(* PLC project Gaia V6.project, CODESYS CODESYS V3.5 SP22 Patch 2 *)
(* stored: creationDateTime 2026-10-21T15:12:01.6200674, modificationDateTime 2026-10-21T14:27:21.3389871 *)

TYPE DUT_EXC_DOSENSOR : STRUCT
  EXC_OUTPUT_SIGNAL : REAL;  (* [EXC : to other equipment] Dissolved oxygen measure *)
  UPI_INPUT_GLOBAL_LOCAL_FUXA : BOOL;  (* [UPI : functional units to equipment] From UPI_LOCAL_FUXA : global FUXA local active *)
  UPI_INPUT_GLOBAL_LOCAL_HMI : BOOL;  (* From UPI_LOCAL_HMI : global HMI local active *)
  UPI_INPUT_GLOBAL_LOCAL_WEBVISU : BOOL;  (* From UPI_LOCAL_webvisu : global HMI local active *)
END_STRUCT;
END_TYPE

TYPE DUT_INT_DIP1500 : STRUCT
  FUXA_LOCAL_REQUEST : BOOL;  (* [Control mode] From FUXA : local request (pulse or maintained) *)
  FUXA_AUTO_REQUEST : BOOL;  (* From FUXA : auto request, releases the individual FUXA local *)
  HMI_LOCAL_REQUEST : BOOL;  (* From HMI : local request (pulse or maintained) *)
  HMI_AUTO_REQUEST : BOOL;  (* From HMI : auto request, releases the individual HMI local *)
  GLOBAL_LOCAL_FUXA : BOOL;  (* From UPI_LOCAL_FUXA : global FUXA local active *)
  GLOBAL_LOCAL_HMI : BOOL;  (* From UPI_LOCAL_HMI : global HMI local active *)
  LOCAL_FUXA_INDIVIDUAL : BOOL;  (* Memory : individual FUXA local, set by local request, reset by auto request *)
  LOCAL_HMI_INDIVIDUAL : BOOL;  (* Memory : individual HMI local, set by local request, reset by auto request *)
  LOCAL_HMI : BOOL;  (* Result : equipment in HMI local (individual or global), unless WEBVISU local is active *)
  LOCAL_FUXA : BOOL;  (* Result : equipment in FUXA local (individual or global), unless WEBVISU or HMI local is active *)
  AUTO : BOOL;  (* Result : no local mode, commands come from the functional units (UPI) *)
  CMD_RUN : BOOL;  (* [Commands (to pump), from the active source] 0 stop, 1 start *)
  CMD_CLOCKWISE : BOOL;  (* 0 counterclockwise, 1 clockwise *)
  CMD_SAVE_FLASH : BOOL;  (* 1 s pulse to coil 0x0003, saves pump parameters to flash *)
  CMD_VOLUME_MODE : BOOL;  (* 0 time mode, 1 volume mode *)
  CMD_SPEED : REAL;  (* rpm *)
  CMD_MAX_SPEED : REAL;  (* rpm *)
  CMD_RUN_SETPOINT : REAL;  (* ms (time mode) or ml (volume mode), 0 = continuous *)
  CMD_CALIB_COEF : REAL;  (* ml/min or rpm *)
  CMD_FOOT_MODE : WORD;  (* Foot switch input mode *)
  CMD_LEVEL_MODE : WORD;  (* Liquid level input mode *)
  CMD_STATE_OUT_MODE : WORD;  (* State output mode *)
  CMD_ADDRESS : WORD;  (* Modbus address *)
  CMD_BAUD_INDEX : WORD;  (* 0=1200 .. 3=9600 .. 7=115200 *)
  PARAM_WRITE_ENABLE : BOOL;  (* [Parameter writing] 1 = write configuration to the pump, 0 = stop writing *)
  FLASH_SAVE_REQUEST : BOOL;  (* Flash save request (rising edge used) *)
  PARAM_VALID : BOOL;  (* Address 1..31, baud index 0..7, max speed > 0, calibration coefficient > 0 *)
  PULSE_500MS : BOOL;  (* [Write triggers] Square wave, 500 ms period, source of the trigger edges *)
  CMD_CHANGED : BOOL;  (* A command value changed this cycle *)
  CMD_WINDOW : BOOL;  (* Command write window, 3 s after the last change *)
  CMD_TRIGGER : BOOL;  (* Command channel trigger *)
  CONFIG_TRIGGER : BOOL;  (* Configuration channel trigger *)
  PREV_RUN : BOOL;  (* [Previous command values] Previous values for change detection *)
  PREV_CLOCKWISE : BOOL;
  PREV_VOLUME_MODE : BOOL;
  PREV_SAVE_FLASH : BOOL;
  PREV_SPEED : REAL;
  PREV_MAX_SPEED : REAL;
  PREV_RUN_SETPOINT : REAL;
  FBK_FIRMWARE_VERSION : WORD;  (* [Feedback (from pump)] 3+5+8 bits (major+minor+revision) *)
  FBK_HARDWARE_VERSION : WORD;  (* 3+5+8 bits (major+sub+reserved) *)
  FBK_TEMPERATURE : WORD;  (* (raw - 500) / 10 = degC, 65535 = not connected *)
  FBK_LEVEL_ALARM : WORD;  (* 0 no alarm, 1 alarm, 65535 = not connected *)
  FBK_DIGITAL_OUTPUT : WORD;  (* Digital output value *)
  FBK_RUN_ACTUAL : REAL;  (* Current run, ms (time mode) or ml (volume mode) *)
  FBK_RUN_TOTAL : REAL;  (* Accumulated run, ms (time mode) or ml (volume mode) *)
  UDINT_TEMP : UDINT;  (* [Work] Work variable, time mode conversion *)
  WEBVISU_LOCAL_REQUEST : BOOL;  (* From WEBVISU : individual local request *)
  WEBVISU_AUTO_REQUEST : BOOL;  (* From WEBVISU : releases individual WEBVISU local (auto wins) *)
  GLOBAL_LOCAL_WEBVISU : BOOL;  (* From UPI_LOCAL_WEBVISU : global local request *)
  LOCAL_WEBVISU_INDIVIDUAL : BOOL;  (* Memory : individual WEBVISU local request *)
  LOCAL_WEBVISU : BOOL;  (* Effective WEBVISU local : highest source priority *)
  SRC_MAX_MOTOR_SPEED : REAL;  (* [Parameter source] Value typed in the active local supervision *)
  SRC_CALIBRATION_COEFFICIENT : REAL;
  SRC_FOOT_SWITCH_INPUT_MODE : WORD;
  SRC_LIQUID_LEVEL_INPUT_MODE : WORD;
  SRC_STATE_OUTPUT_MODE : WORD;
  SRC_COMMUNICATION_ADDRESS : WORD;
  SRC_BAUD_RATE_INDEX : WORD;
  PREV_SRC_MAX_MOTOR_SPEED : REAL;  (* [Parameter change detection] Previous source values *)
  PREV_SRC_CALIBRATION_COEFFICIENT : REAL;
  PREV_SRC_FOOT_SWITCH_INPUT_MODE : WORD;
  PREV_SRC_LIQUID_LEVEL_INPUT_MODE : WORD;
  PREV_SRC_STATE_OUTPUT_MODE : WORD;
  PREV_SRC_COMMUNICATION_ADDRESS : WORD;
  PREV_SRC_BAUD_RATE_INDEX : WORD;
  PREV_LOCAL_WEBVISU : BOOL;  (* Previous control mode, to ignore the cycle where the source changes *)
  PREV_LOCAL_HMI : BOOL;
  PREV_LOCAL_FUXA : BOOL;
  SOURCE_CHANGED : BOOL;  (* The active local source changed this cycle : no parameter is taken *)
END_STRUCT;
END_TYPE

TYPE DUT_IO_DOSENSOR : STRUCT
  INPUT_SIGNAL : DWORD;  (* [INPUT (field to PLC)] Analog input, raw value *)
  INPUT_SENSOR_FAULT : BOOL;  (* Digital input, sensor fault *)
  OUTPUT_CALIBRATION_HIGH : BOOL;  (* [OUTPUT (PLC to field)] Digital output, high calibration *)
  OUTPUT_CALIBRATION_LOW : BOOL;  (* Digital output, low calibration *)
END_STRUCT;
END_TYPE

TYPE DUT_INT_DOSENSOR : STRUCT
  FUXA_LOCAL_REQUEST : BOOL;  (* [Control mode] From FUXA : local request (pulse or maintained) *)
  FUXA_AUTO_REQUEST : BOOL;  (* From FUXA : auto request, releases the individual FUXA local *)
  HMI_LOCAL_REQUEST : BOOL;  (* From HMI : local request (pulse or maintained) *)
  HMI_AUTO_REQUEST : BOOL;  (* From HMI : auto request, releases the individual HMI local *)
  GLOBAL_LOCAL_FUXA : BOOL;  (* From UPI_LOCAL_FUXA : global FUXA local active *)
  GLOBAL_LOCAL_HMI : BOOL;  (* From UPI_LOCAL_HMI : global HMI local active *)
  LOCAL_FUXA_INDIVIDUAL : BOOL;  (* Memory : individual FUXA local, set by local request, reset by auto request *)
  LOCAL_HMI_INDIVIDUAL : BOOL;  (* Memory : individual HMI local, set by local request, reset by auto request *)
  LOCAL_HMI : BOOL;  (* Result : equipment in HMI local (individual or global), unless WEBVISU local is active *)
  LOCAL_FUXA : BOOL;  (* Result : equipment in FUXA local (individual or global), unless WEBVISU or HMI local is active *)
  WEBVISU_LOCAL_REQUEST : BOOL;  (* From WEBVISU : local request (pulse or maintained) *)
  WEBVISU_AUTO_REQUEST : BOOL;  (* From WEBVISU : auto request, releases the individual WEBVISU local *)
  LOCAL_WEBVISU_INDIVIDUAL : BOOL;  (* Memory : individual WEBVISU local, set by local request, reset by auto request *)
  LOCAL_WEBVISU : BOOL;  (* Result : equipment in WEBVISU local (individual or global), has priority *)
  AUTO : BOOL;  (* Result : no local mode, commands come from the functional units (UPI) *)
  SIGNAL_RAW : DWORD;  (* [Inputs] Raw analog input *)
  FAULT : BOOL;  (* Sensor fault (digital input) *)
  CALIB_HIGH_REQUEST : BOOL;  (* High calibration request from the active source *)
  CALIB_LOW_REQUEST : BOOL;  (* Low calibration request from the active source *)
  SIGNAL : REAL;  (* [Results] Scaled measure *)
  CALIB_HIGH : BOOL;  (* High calibration pulse to sensor (1 s) *)
  CALIB_LOW : BOOL;  (* Low calibration pulse to sensor (1 s) *)
  CALIB_DONE : BOOL;  (* Calibration done message (5 s) *)
  GLOBAL_LOCAL_WEBVISU : BOOL;  (* From UPI_LOCAL_WEBVISU : global local request *)
END_STRUCT;
END_TYPE

TYPE DUT_COM_DOSENSOR : STRUCT
  SCADA_INPUT_CALIBRATION_HIGH : BOOL;  (* [SCADA (FUXA) : input (to PLC)] Coil 1 | DO Calibration High *)
  SCADA_INPUT_CALIBRATION_LOW : BOOL;  (* Coil 2 | DO Calibration Low *)
  SCADA_INPUT_LOCAL_REQUEST : BOOL;  (* Coil 8 | DO Sensor Local Request *)
  SCADA_INPUT_AUTO_REQUEST : BOOL;  (* Coil 9 | DO Sensor Auto Request *)
  SCADA_OUTPUT_FAULT : BOOL;  (* [SCADA (FUXA) : output (from PLC)] DI 10001 | Do sensor fault *)
  SCADA_OUTPUT_CALIBRATION_DONE : BOOL;  (* DI 10002 | Do sensor calibration done *)
  SCADA_OUTPUT_LOCAL_FUXA_ACTIVE : BOOL;  (* DI 10013 | DO Sensor Local FUXA Active *)
  SCADA_OUTPUT_LOCAL_HMI_ACTIVE : BOOL;  (* DI 10014 | DO Sensor Local HMI Active *)
  SCADA_OUTPUT_SIGNAL : DUT_Union_Real_Word;  (* IR 89-90 | DO Sensor Signal *)
  HMI_INPUT_CALIBRATION_HIGH : BOOL;  (* [HMI (local panel, FUXA address + 1000) : input (to PLC)] Coil 1001 | DO Calibration High *)
  HMI_INPUT_CALIBRATION_LOW : BOOL;  (* Coil 1002 | DO Calibration Low *)
  HMI_INPUT_LOCAL_REQUEST : BOOL;  (* Coil 1008 | DO Sensor Local Request *)
  HMI_INPUT_AUTO_REQUEST : BOOL;  (* Coil 1009 | DO Sensor Auto Request *)
  HMI_OUTPUT_FAULT : BOOL;  (* [HMI (local panel, FUXA address + 1000) : output (from PLC)] DI 11001 | Do sensor fault *)
  HMI_OUTPUT_CALIBRATION_DONE : BOOL;  (* DI 11002 | Do sensor calibration done *)
  HMI_OUTPUT_LOCAL_ACTIVE : BOOL;  (* DI 11014 | DO Sensor Local Active *)
  HMI_OUTPUT_SIGNAL : DUT_Union_Real_Word;  (* IR 1089-1090 | DO Sensor Signal *)
  WEBVISU_INPUT_CALIBRATION_HIGH : BOOL;  (* DO Calibration High *)
  WEBVISU_INPUT_CALIBRATION_LOW : BOOL;  (* DO Calibration Low *)
  WEBVISU_INPUT_LOCAL_REQUEST : BOOL;  (* DO Sensor Local Request *)
  WEBVISU_INPUT_AUTO_REQUEST : BOOL;  (* DO Sensor Auto Request *)
  WEBVISU_OUTPUT_FAULT : BOOL;  (* Do sensor fault *)
  WEBVISU_OUTPUT_CALIBRATION_DONE : BOOL;  (* Do sensor calibration done *)
  WEBVISU_OUTPUT_LOCAL_ACTIVE : BOOL;  (* DO Sensor Local Active *)
  WEBVISU_OUTPUT_SIGNAL : DUT_Union_Real_Word;  (* DO Sensor Signal *)
  WEBVISU_OUTPUT_LOCAL_FUXA_ACTIVE : BOOL;  (* Effective FUXA local mode (masked by WEBVISU and HMI priority) *)
  WEBVISU_OUTPUT_LOCAL_HMI_ACTIVE : BOOL;  (* Effective HMI local mode (masked by WEBVISU priority) *)
END_STRUCT;
END_TYPE

TYPE DUT_INT_ADM100W : STRUCT
  FUXA_LOCAL_REQUEST : BOOL;  (* [Control mode] From FUXA : local request (pulse or maintained) *)
  FUXA_AUTO_REQUEST : BOOL;  (* From FUXA : auto request, releases the individual FUXA local *)
  HMI_LOCAL_REQUEST : BOOL;  (* From HMI : local request (pulse or maintained) *)
  HMI_AUTO_REQUEST : BOOL;  (* From HMI : auto request, releases the individual HMI local *)
  GLOBAL_LOCAL_FUXA : BOOL;  (* From UPI_LOCAL_FUXA : global FUXA local active *)
  GLOBAL_LOCAL_HMI : BOOL;  (* From UPI_LOCAL_HMI : global HMI local active *)
  LOCAL_FUXA_INDIVIDUAL : BOOL;  (* Memory : individual FUXA local, set by local request, reset by auto request *)
  LOCAL_HMI_INDIVIDUAL : BOOL;  (* Memory : individual HMI local, set by local request, reset by auto request *)
  LOCAL_HMI : BOOL;  (* Result : equipment in HMI local (individual or global), unless WEBVISU local is active *)
  LOCAL_FUXA : BOOL;  (* Result : equipment in FUXA local (individual or global), unless WEBVISU or HMI local is active *)
  AUTO : BOOL;  (* Result : no local mode, commands come from the functional units (UPI) *)
  ALARM_1 : BOOL;  (* [Alarms] Alarm 1 status *)
  ALARM_2 : BOOL;  (* Alarm 2 status *)
  ALARM_3 : BOOL;  (* Alarm 3 status *)
  ALARM_4 : BOOL;  (* Alarm 4 status *)
  ALARM_5 : BOOL;  (* Alarm 5 status *)
  ALARM_6 : BOOL;  (* Alarm 6 status *)
  ALARM_7 : BOOL;  (* Alarm 7 status *)
  ALARM_8 : BOOL;  (* Alarm 8 status *)
  ALARM_9 : BOOL;  (* Alarm 9 status *)
  ALARM_10 : BOOL;  (* Alarm 10 status *)
  FREQUENCY : REAL;  (* [Measures] Frequency | Hz *)
  L1_L2_VOLTAGE : REAL;  (* L1-L2 Voltage | V *)
  L1_N_VOLTAGE : REAL;  (* L1-N Voltage | V *)
  L1_CURRENT : REAL;  (* L1 Current | A *)
  L1_ACTIVE_POWER : REAL;  (* L1 Active Power | W *)
  L1_APPARENT_POWER : REAL;  (* L1 Apparent Power | VA *)
  L1_REACTIVE_POWER : REAL;  (* L1 Reactive Power | W *)
  L1_CURRENT_PHASE_ANGLE : REAL;  (* L1 Current Phase Angle | deg *)
  L1_POWER_FACTOR : REAL;  (* L1 Power Factor | - *)
  L1_VOLTAGE_THD : REAL;  (* L1 Voltage THD | % *)
  L1_CURRENT_THD : REAL;  (* L1 Current THD | % *)
  L1_MAX_LOAD : REAL;  (* L1 Max Load | % of 60 A *)
  L1_L2_VOLTAGE_PHASE_ANGLE : REAL;  (* L1-L2 Voltage Phase Angle | deg *)
  L2_L3_VOLTAGE : REAL;  (* L2-L3 Voltage | V *)
  L2_N_VOLTAGE : REAL;  (* L2-N Voltage | V *)
  L2_CURRENT : REAL;  (* L2 Current | A *)
  L2_ACTIVE_POWER : REAL;  (* L2 Active Power | W *)
  L2_APPARENT_POWER : REAL;  (* L2 Apparent Power | VA *)
  L2_REACTIVE_POWER : REAL;  (* L2 Reactive Power | W *)
  L2_CURRENT_PHASE_ANGLE : REAL;  (* L2 Current Phase Angle | deg *)
  L2_POWER_FACTOR : REAL;  (* L2 Power Factor | - *)
  L2_VOLTAGE_THD : REAL;  (* L2 Voltage THD | % *)
  L2_CURRENT_THD : REAL;  (* L2 Current THD | % *)
  L2_MAX_LOAD : REAL;  (* L2 Max Load | % of 60 A *)
  L1_L3_VOLTAGE_PHASE_ANGLE : REAL;  (* L1-L3 Voltage Phase Angle | deg *)
  L3_L1_VOLTAGE : REAL;  (* L3-L1 Voltage | V *)
  L3_N_VOLTAGE : REAL;  (* L3-N Voltage | V *)
  L3_CURRENT : REAL;  (* L3 Current | A *)
  L3_ACTIVE_POWER : REAL;  (* L3 Active Power | W *)
  L3_APPARENT_POWER : REAL;  (* L3 Apparent Power | VA *)
  L3_REACTIVE_POWER : REAL;  (* L3 Reactive Power | W *)
  L3_CURRENT_PHASE_ANGLE : REAL;  (* L3 Current Phase Angle | deg *)
  L3_POWER_FACTOR : REAL;  (* L3 Power Factor | - *)
  L3_VOLTAGE_THD : REAL;  (* L3 Voltage THD | % *)
  L3_CURRENT_THD : REAL;  (* L3 Current THD | % *)
  L3_MAX_LOAD : REAL;  (* L3 Max Load | % of 60 A *)
  INTERNAL_TEMPERATURE : REAL;  (* Internal Temperature | degC *)
  ACTIVE_ENERGY : REAL;  (* Active Energy | kWh *)
  APPARENT_ENERGY : REAL;  (* Apparent Energy | per ADM100W config *)
  REACTIVE_ENERGY : REAL;  (* Reactive Energy | kWh *)
  TOTAL_ACTIVE_POWER : REAL;  (* Total Active Power | W *)
  TOTAL_APPARENT_POWER : REAL;  (* Total Apparent Power | VA *)
  TOTAL_REACTIVE_POWER : REAL;  (* Total Reactive Power | W *)
  ALL_PHASE_POWER_FACTOR : REAL;  (* All Phase Power Factor | - *)
  WEBVISU_LOCAL_REQUEST : BOOL;  (* From WEBVISU : individual local request *)
  WEBVISU_AUTO_REQUEST : BOOL;  (* From WEBVISU : releases individual WEBVISU local (auto wins) *)
  GLOBAL_LOCAL_WEBVISU : BOOL;  (* From UPI_LOCAL_WEBVISU : global local request *)
  LOCAL_WEBVISU_INDIVIDUAL : BOOL;  (* Memory : individual WEBVISU local request *)
  LOCAL_WEBVISU : BOOL;  (* Effective WEBVISU local : highest source priority *)
END_STRUCT;
END_TYPE

TYPE DUT_COM_UPI_LOCAL_FUXA : STRUCT
  SCADA_INPUT_LOCAL_REQUEST : BOOL;  (* [SCADA (FUXA) : input (to PLC)] Coil 14 | Global Local FUXA Request *)
  SCADA_INPUT_AUTO_REQUEST : BOOL;  (* Coil 15 | Global Auto FUXA Request *)
  SCADA_OUTPUT_LOCAL_ACTIVE : BOOL;  (* [SCADA (FUXA) : output (from PLC)] DI 10019 | Global Local FUXA Active *)
END_STRUCT;
END_TYPE

TYPE DUT_IO_ADM100W : STRUCT
  SPARE : BOOL;  (* Placeholder, structure not used yet *)
END_STRUCT;
END_TYPE

TYPE DUT_COM_ADM100W : STRUCT
  COM_INPUT_IR : ARRAY[0..87] OF WORD;  (* [COM : Modbus RTU, input (equipment to PLC)] Input registers 0..87, 32-bit float, MSW first (ABCD) *)
  COM_INPUT_COILS : ARRAY[0..1] OF BYTE;  (* Coils 0..9 = alarms 1..10 (byte.bit) *)
  SCADA_INPUT_LOCAL_REQUEST : BOOL;  (* [SCADA (FUXA) : input (to PLC)] Coil 12 | ADM100W Local Request *)
  SCADA_INPUT_AUTO_REQUEST : BOOL;  (* Coil 13 | ADM100W Auto Request *)
  SCADA_OUTPUT_ALARM_1_STATUS : BOOL;  (* [SCADA (FUXA) : output (from PLC)] DI 10003 | ADM100W Alarm 1 Status *)
  SCADA_OUTPUT_ALARM_2_STATUS : BOOL;  (* DI 10004 | ADM100W Alarm 2 Status *)
  SCADA_OUTPUT_ALARM_3_STATUS : BOOL;  (* DI 10005 | ADM100W Alarm 3 Status *)
  SCADA_OUTPUT_ALARM_4_STATUS : BOOL;  (* DI 10006 | ADM100W Alarm 4 Status *)
  SCADA_OUTPUT_ALARM_5_STATUS : BOOL;  (* DI 10007 | ADM100W Alarm 5 Status *)
  SCADA_OUTPUT_ALARM_6_STATUS : BOOL;  (* DI 10008 | ADM100W Alarm 6 Status *)
  SCADA_OUTPUT_ALARM_7_STATUS : BOOL;  (* DI 10009 | ADM100W Alarm 7 Status *)
  SCADA_OUTPUT_ALARM_8_STATUS : BOOL;  (* DI 10010 | ADM100W Alarm 8 Status *)
  SCADA_OUTPUT_ALARM_9_STATUS : BOOL;  (* DI 10011 | ADM100W Alarm 9 Status *)
  SCADA_OUTPUT_ALARM_10_STATUS : BOOL;  (* DI 10012 | ADM100W Alarm 10 Status *)
  SCADA_OUTPUT_LOCAL_FUXA_ACTIVE : BOOL;  (* DI 10017 | ADM100W Local FUXA Active *)
  SCADA_OUTPUT_LOCAL_HMI_ACTIVE : BOOL;  (* DI 10018 | ADM100W Local HMI Active *)
  SCADA_OUTPUT_FREQUENCY : DUT_Union_Real_Word;  (* IR 1-2 | ADM100W Frequency | Hz *)
  SCADA_OUTPUT_L1_L2_VOLTAGE : DUT_Union_Real_Word;  (* IR 3-4 | ADM100W L1-L2 Voltage | V *)
  SCADA_OUTPUT_L1_N_VOLTAGE : DUT_Union_Real_Word;  (* IR 5-6 | ADM100W L1-N Voltage | V *)
  SCADA_OUTPUT_L1_CURRENT : DUT_Union_Real_Word;  (* IR 7-8 | ADM100W L1 Current | A *)
  SCADA_OUTPUT_L1_ACTIVE_POWER : DUT_Union_Real_Word;  (* IR 9-10 | ADM100W L1 Active Power *)
  SCADA_OUTPUT_L1_APPARENT_POWER : DUT_Union_Real_Word;  (* IR 11-12 | ADM100W L1 Apparent Power *)
  SCADA_OUTPUT_L1_REACTIVE_POWER : DUT_Union_Real_Word;  (* IR 13-14 | ADM100W L1 Reactive Power *)
  SCADA_OUTPUT_L1_CURRENT_PHASE_ANGLE : DUT_Union_Real_Word;  (* IR 15-16 | ADM100W L1 Current Phase Angle | deg *)
  SCADA_OUTPUT_L1_POWER_FACTOR : DUT_Union_Real_Word;  (* IR 17-18 | ADM100W L1 Power Factor *)
  SCADA_OUTPUT_L1_VOLTAGE_THD : DUT_Union_Real_Word;  (* IR 19-20 | ADM100W L1 Voltage THD | % *)
  SCADA_OUTPUT_L1_CURRENT_THD : DUT_Union_Real_Word;  (* IR 21-22 | ADM100W L1 Current THD | % *)
  SCADA_OUTPUT_L1_MAX_LOAD : DUT_Union_Real_Word;  (* IR 23-24 | ADM100W L1 Max Load *)
  SCADA_OUTPUT_L1_L2_VOLTAGE_PHASE_ANGLE : DUT_Union_Real_Word;  (* IR 25-26 | ADM100W L1-L2 Voltage Phase Angle | deg *)
  SCADA_OUTPUT_L2_L3_VOLTAGE : DUT_Union_Real_Word;  (* IR 27-28 | ADM100W L2-L3 Voltage | V *)
  SCADA_OUTPUT_L2_N_VOLTAGE : DUT_Union_Real_Word;  (* IR 29-30 | ADM100W L2-N Voltage | V *)
  SCADA_OUTPUT_L2_CURRENT : DUT_Union_Real_Word;  (* IR 31-32 | ADM100W L2 Current | A *)
  SCADA_OUTPUT_L2_ACTIVE_POWER : DUT_Union_Real_Word;  (* IR 33-34 | ADM100W L2 Active Power *)
  SCADA_OUTPUT_L2_APPARENT_POWER : DUT_Union_Real_Word;  (* IR 35-36 | ADM100W L2 Apparent Power *)
  SCADA_OUTPUT_L2_REACTIVE_POWER : DUT_Union_Real_Word;  (* IR 37-38 | ADM100W L2 Reactive Power *)
  SCADA_OUTPUT_L2_CURRENT_PHASE_ANGLE : DUT_Union_Real_Word;  (* IR 39-40 | ADM100W L2 Current Phase Angle | deg *)
  SCADA_OUTPUT_L2_POWER_FACTOR : DUT_Union_Real_Word;  (* IR 41-42 | ADM100W L2 Power Factor *)
  SCADA_OUTPUT_L2_VOLTAGE_THD : DUT_Union_Real_Word;  (* IR 43-44 | ADM100W L2 Voltage THD | % *)
  SCADA_OUTPUT_L2_CURRENT_THD : DUT_Union_Real_Word;  (* IR 45-46 | ADM100W L2 Current THD | % *)
  SCADA_OUTPUT_L2_MAX_LOAD : DUT_Union_Real_Word;  (* IR 47-48 | ADM100W L2 Max Load *)
  SCADA_OUTPUT_L1_L3_VOLTAGE_PHASE_ANGLE : DUT_Union_Real_Word;  (* IR 49-50 | ADM100W L1-L3 Voltage Phase Angle | deg *)
  SCADA_OUTPUT_L3_L1_VOLTAGE : DUT_Union_Real_Word;  (* IR 51-52 | ADM100W L3-L1 Voltage | V *)
  SCADA_OUTPUT_L3_N_VOLTAGE : DUT_Union_Real_Word;  (* IR 53-54 | ADM100W L3-N Voltage | V *)
  SCADA_OUTPUT_L3_CURRENT : DUT_Union_Real_Word;  (* IR 55-56 | ADM100W L3 Current | A *)
  SCADA_OUTPUT_L3_ACTIVE_POWER : DUT_Union_Real_Word;  (* IR 57-58 | ADM100W L3 Active Power *)
  SCADA_OUTPUT_L3_APPARENT_POWER : DUT_Union_Real_Word;  (* IR 59-60 | ADM100W L3 Apparent Power *)
  SCADA_OUTPUT_L3_REACTIVE_POWER : DUT_Union_Real_Word;  (* IR 61-62 | ADM100W L3 Reactive Power *)
  SCADA_OUTPUT_L3_CURRENT_PHASE_ANGLE : DUT_Union_Real_Word;  (* IR 63-64 | ADM100W L3 Current Phase Angle | deg *)
  SCADA_OUTPUT_L3_POWER_FACTOR : DUT_Union_Real_Word;  (* IR 65-66 | ADM100W L3 Power Factor *)
  SCADA_OUTPUT_L3_VOLTAGE_THD : DUT_Union_Real_Word;  (* IR 67-68 | ADM100W L3 Voltage THD | % *)
  SCADA_OUTPUT_L3_CURRENT_THD : DUT_Union_Real_Word;  (* IR 69-70 | ADM100W L3 Current THD | % *)
  SCADA_OUTPUT_L3_MAX_LOAD : DUT_Union_Real_Word;  (* IR 71-72 | ADM100W L3 Max Load *)
  SCADA_OUTPUT_INTERNAL_TEMPERATURE : DUT_Union_Real_Word;  (* IR 73-74 | ADM100W Internal Temperature *)
  SCADA_OUTPUT_ACTIVE_ENERGY : DUT_Union_Real_Word;  (* IR 75-76 | ADM100W Active Energy *)
  SCADA_OUTPUT_APPARENT_ENERGY : DUT_Union_Real_Word;  (* IR 77-78 | ADM100W Apparent Energy *)
  SCADA_OUTPUT_REACTIVE_ENERGY : DUT_Union_Real_Word;  (* IR 79-80 | ADM100W Reactive Energy *)
  SCADA_OUTPUT_TOTAL_ACTIVE_POWER : DUT_Union_Real_Word;  (* IR 81-82 | ADM100W Total Active Power *)
  SCADA_OUTPUT_TOTAL_APPARENT_POWER : DUT_Union_Real_Word;  (* IR 83-84 | ADM100W Total Apparent Power *)
  SCADA_OUTPUT_TOTAL_REACTIVE_POWER : DUT_Union_Real_Word;  (* IR 85-86 | ADM100W Total Reactive Power *)
  SCADA_OUTPUT_ALL_PHASE_POWER_FACTOR : DUT_Union_Real_Word;  (* IR 87-88 | ADM100W All Phase Power Factor *)
  HMI_INPUT_LOCAL_REQUEST : BOOL;  (* [HMI (local panel, FUXA address + 1000) : input (to PLC)] Coil 1012 | ADM100W Local Request *)
  HMI_INPUT_AUTO_REQUEST : BOOL;  (* Coil 1013 | ADM100W Auto Request *)
  HMI_OUTPUT_ALARM_1_STATUS : BOOL;  (* [HMI (local panel, FUXA address + 1000) : output (from PLC)] DI 11003 | ADM100W Alarm 1 Status *)
  HMI_OUTPUT_ALARM_2_STATUS : BOOL;  (* DI 11004 | ADM100W Alarm 2 Status *)
  HMI_OUTPUT_ALARM_3_STATUS : BOOL;  (* DI 11005 | ADM100W Alarm 3 Status *)
  HMI_OUTPUT_ALARM_4_STATUS : BOOL;  (* DI 11006 | ADM100W Alarm 4 Status *)
  HMI_OUTPUT_ALARM_5_STATUS : BOOL;  (* DI 11007 | ADM100W Alarm 5 Status *)
  HMI_OUTPUT_ALARM_6_STATUS : BOOL;  (* DI 11008 | ADM100W Alarm 6 Status *)
  HMI_OUTPUT_ALARM_7_STATUS : BOOL;  (* DI 11009 | ADM100W Alarm 7 Status *)
  HMI_OUTPUT_ALARM_8_STATUS : BOOL;  (* DI 11010 | ADM100W Alarm 8 Status *)
  HMI_OUTPUT_ALARM_9_STATUS : BOOL;  (* DI 11011 | ADM100W Alarm 9 Status *)
  HMI_OUTPUT_ALARM_10_STATUS : BOOL;  (* DI 11012 | ADM100W Alarm 10 Status *)
  HMI_OUTPUT_LOCAL_ACTIVE : BOOL;  (* DI 11018 | ADM100W Local Active *)
  HMI_OUTPUT_FREQUENCY : DUT_Union_Real_Word;  (* IR 1001-1002 | ADM100W Frequency | Hz *)
  HMI_OUTPUT_L1_L2_VOLTAGE : DUT_Union_Real_Word;  (* IR 1003-1004 | ADM100W L1-L2 Voltage | V *)
  HMI_OUTPUT_L1_N_VOLTAGE : DUT_Union_Real_Word;  (* IR 1005-1006 | ADM100W L1-N Voltage | V *)
  HMI_OUTPUT_L1_CURRENT : DUT_Union_Real_Word;  (* IR 1007-1008 | ADM100W L1 Current | A *)
  HMI_OUTPUT_L1_ACTIVE_POWER : DUT_Union_Real_Word;  (* IR 1009-1010 | ADM100W L1 Active Power *)
  HMI_OUTPUT_L1_APPARENT_POWER : DUT_Union_Real_Word;  (* IR 1011-1012 | ADM100W L1 Apparent Power *)
  HMI_OUTPUT_L1_REACTIVE_POWER : DUT_Union_Real_Word;  (* IR 1013-1014 | ADM100W L1 Reactive Power *)
  HMI_OUTPUT_L1_CURRENT_PHASE_ANGLE : DUT_Union_Real_Word;  (* IR 1015-1016 | ADM100W L1 Current Phase Angle | deg *)
  HMI_OUTPUT_L1_POWER_FACTOR : DUT_Union_Real_Word;  (* IR 1017-1018 | ADM100W L1 Power Factor *)
  HMI_OUTPUT_L1_VOLTAGE_THD : DUT_Union_Real_Word;  (* IR 1019-1020 | ADM100W L1 Voltage THD | % *)
  HMI_OUTPUT_L1_CURRENT_THD : DUT_Union_Real_Word;  (* IR 1021-1022 | ADM100W L1 Current THD | % *)
  HMI_OUTPUT_L1_MAX_LOAD : DUT_Union_Real_Word;  (* IR 1023-1024 | ADM100W L1 Max Load *)
  HMI_OUTPUT_L1_L2_VOLTAGE_PHASE_ANGLE : DUT_Union_Real_Word;  (* IR 1025-1026 | ADM100W L1-L2 Voltage Phase Angle | deg *)
  HMI_OUTPUT_L2_L3_VOLTAGE : DUT_Union_Real_Word;  (* IR 1027-1028 | ADM100W L2-L3 Voltage | V *)
  HMI_OUTPUT_L2_N_VOLTAGE : DUT_Union_Real_Word;  (* IR 1029-1030 | ADM100W L2-N Voltage | V *)
  HMI_OUTPUT_L2_CURRENT : DUT_Union_Real_Word;  (* IR 1031-1032 | ADM100W L2 Current | A *)
  HMI_OUTPUT_L2_ACTIVE_POWER : DUT_Union_Real_Word;  (* IR 1033-1034 | ADM100W L2 Active Power *)
  HMI_OUTPUT_L2_APPARENT_POWER : DUT_Union_Real_Word;  (* IR 1035-1036 | ADM100W L2 Apparent Power *)
  HMI_OUTPUT_L2_REACTIVE_POWER : DUT_Union_Real_Word;  (* IR 1037-1038 | ADM100W L2 Reactive Power *)
  HMI_OUTPUT_L2_CURRENT_PHASE_ANGLE : DUT_Union_Real_Word;  (* IR 1039-1040 | ADM100W L2 Current Phase Angle | deg *)
  HMI_OUTPUT_L2_POWER_FACTOR : DUT_Union_Real_Word;  (* IR 1041-1042 | ADM100W L2 Power Factor *)
  HMI_OUTPUT_L2_VOLTAGE_THD : DUT_Union_Real_Word;  (* IR 1043-1044 | ADM100W L2 Voltage THD | % *)
  HMI_OUTPUT_L2_CURRENT_THD : DUT_Union_Real_Word;  (* IR 1045-1046 | ADM100W L2 Current THD | % *)
  HMI_OUTPUT_L2_MAX_LOAD : DUT_Union_Real_Word;  (* IR 1047-1048 | ADM100W L2 Max Load *)
  HMI_OUTPUT_L1_L3_VOLTAGE_PHASE_ANGLE : DUT_Union_Real_Word;  (* IR 1049-1050 | ADM100W L1-L3 Voltage Phase Angle | deg *)
  HMI_OUTPUT_L3_L1_VOLTAGE : DUT_Union_Real_Word;  (* IR 1051-1052 | ADM100W L3-L1 Voltage | V *)
  HMI_OUTPUT_L3_N_VOLTAGE : DUT_Union_Real_Word;  (* IR 1053-1054 | ADM100W L3-N Voltage | V *)
  HMI_OUTPUT_L3_CURRENT : DUT_Union_Real_Word;  (* IR 1055-1056 | ADM100W L3 Current | A *)
  HMI_OUTPUT_L3_ACTIVE_POWER : DUT_Union_Real_Word;  (* IR 1057-1058 | ADM100W L3 Active Power *)
  HMI_OUTPUT_L3_APPARENT_POWER : DUT_Union_Real_Word;  (* IR 1059-1060 | ADM100W L3 Apparent Power *)
  HMI_OUTPUT_L3_REACTIVE_POWER : DUT_Union_Real_Word;  (* IR 1061-1062 | ADM100W L3 Reactive Power *)
  HMI_OUTPUT_L3_CURRENT_PHASE_ANGLE : DUT_Union_Real_Word;  (* IR 1063-1064 | ADM100W L3 Current Phase Angle | deg *)
  HMI_OUTPUT_L3_POWER_FACTOR : DUT_Union_Real_Word;  (* IR 1065-1066 | ADM100W L3 Power Factor *)
  HMI_OUTPUT_L3_VOLTAGE_THD : DUT_Union_Real_Word;  (* IR 1067-1068 | ADM100W L3 Voltage THD | % *)
  HMI_OUTPUT_L3_CURRENT_THD : DUT_Union_Real_Word;  (* IR 1069-1070 | ADM100W L3 Current THD | % *)
  HMI_OUTPUT_L3_MAX_LOAD : DUT_Union_Real_Word;  (* IR 1071-1072 | ADM100W L3 Max Load *)
  HMI_OUTPUT_INTERNAL_TEMPERATURE : DUT_Union_Real_Word;  (* IR 1073-1074 | ADM100W Internal Temperature *)
  HMI_OUTPUT_ACTIVE_ENERGY : DUT_Union_Real_Word;  (* IR 1075-1076 | ADM100W Active Energy *)
  HMI_OUTPUT_APPARENT_ENERGY : DUT_Union_Real_Word;  (* IR 1077-1078 | ADM100W Apparent Energy *)
  HMI_OUTPUT_REACTIVE_ENERGY : DUT_Union_Real_Word;  (* IR 1079-1080 | ADM100W Reactive Energy *)
  HMI_OUTPUT_TOTAL_ACTIVE_POWER : DUT_Union_Real_Word;  (* IR 1081-1082 | ADM100W Total Active Power *)
  HMI_OUTPUT_TOTAL_APPARENT_POWER : DUT_Union_Real_Word;  (* IR 1083-1084 | ADM100W Total Apparent Power *)
  HMI_OUTPUT_TOTAL_REACTIVE_POWER : DUT_Union_Real_Word;  (* IR 1085-1086 | ADM100W Total Reactive Power *)
  HMI_OUTPUT_ALL_PHASE_POWER_FACTOR : DUT_Union_Real_Word;  (* IR 1087-1088 | ADM100W All Phase Power Factor *)
  WEBVISU_INPUT_LOCAL_REQUEST : BOOL;  (* [WEBVISU : direct IEC variable] ADM100W Local Request *)
  WEBVISU_INPUT_AUTO_REQUEST : BOOL;  (* [WEBVISU : direct IEC variable] ADM100W Auto Request *)
  WEBVISU_OUTPUT_ALARM_1_STATUS : BOOL;  (* [WEBVISU : direct IEC variable] ADM100W Alarm 1 Status *)
  WEBVISU_OUTPUT_ALARM_2_STATUS : BOOL;  (* [WEBVISU : direct IEC variable] ADM100W Alarm 2 Status *)
  WEBVISU_OUTPUT_ALARM_3_STATUS : BOOL;  (* [WEBVISU : direct IEC variable] ADM100W Alarm 3 Status *)
  WEBVISU_OUTPUT_ALARM_4_STATUS : BOOL;  (* [WEBVISU : direct IEC variable] ADM100W Alarm 4 Status *)
  WEBVISU_OUTPUT_ALARM_5_STATUS : BOOL;  (* [WEBVISU : direct IEC variable] ADM100W Alarm 5 Status *)
  WEBVISU_OUTPUT_ALARM_6_STATUS : BOOL;  (* [WEBVISU : direct IEC variable] ADM100W Alarm 6 Status *)
  WEBVISU_OUTPUT_ALARM_7_STATUS : BOOL;  (* [WEBVISU : direct IEC variable] ADM100W Alarm 7 Status *)
  WEBVISU_OUTPUT_ALARM_8_STATUS : BOOL;  (* [WEBVISU : direct IEC variable] ADM100W Alarm 8 Status *)
  WEBVISU_OUTPUT_ALARM_9_STATUS : BOOL;  (* [WEBVISU : direct IEC variable] ADM100W Alarm 9 Status *)
  WEBVISU_OUTPUT_ALARM_10_STATUS : BOOL;  (* [WEBVISU : direct IEC variable] ADM100W Alarm 10 Status *)
  WEBVISU_OUTPUT_LOCAL_ACTIVE : BOOL;  (* [WEBVISU : direct IEC variable] ADM100W Local Active *)
  WEBVISU_OUTPUT_FREQUENCY : DUT_Union_Real_Word;  (* [WEBVISU : direct IEC variable] ADM100W Frequency | Hz *)
  WEBVISU_OUTPUT_L1_L2_VOLTAGE : DUT_Union_Real_Word;  (* [WEBVISU : direct IEC variable] ADM100W L1-L2 Voltage | V *)
  WEBVISU_OUTPUT_L1_N_VOLTAGE : DUT_Union_Real_Word;  (* [WEBVISU : direct IEC variable] ADM100W L1-N Voltage | V *)
  WEBVISU_OUTPUT_L1_CURRENT : DUT_Union_Real_Word;  (* [WEBVISU : direct IEC variable] ADM100W L1 Current | A *)
  WEBVISU_OUTPUT_L1_ACTIVE_POWER : DUT_Union_Real_Word;  (* [WEBVISU : direct IEC variable] ADM100W L1 Active Power *)
  WEBVISU_OUTPUT_L1_APPARENT_POWER : DUT_Union_Real_Word;  (* [WEBVISU : direct IEC variable] ADM100W L1 Apparent Power *)
  WEBVISU_OUTPUT_L1_REACTIVE_POWER : DUT_Union_Real_Word;  (* [WEBVISU : direct IEC variable] ADM100W L1 Reactive Power *)
  WEBVISU_OUTPUT_L1_CURRENT_PHASE_ANGLE : DUT_Union_Real_Word;  (* [WEBVISU : direct IEC variable] ADM100W L1 Current Phase Angle | deg *)
  WEBVISU_OUTPUT_L1_POWER_FACTOR : DUT_Union_Real_Word;  (* [WEBVISU : direct IEC variable] ADM100W L1 Power Factor *)
  WEBVISU_OUTPUT_L1_VOLTAGE_THD : DUT_Union_Real_Word;  (* [WEBVISU : direct IEC variable] ADM100W L1 Voltage THD | % *)
  WEBVISU_OUTPUT_L1_CURRENT_THD : DUT_Union_Real_Word;  (* [WEBVISU : direct IEC variable] ADM100W L1 Current THD | % *)
  WEBVISU_OUTPUT_L1_MAX_LOAD : DUT_Union_Real_Word;  (* [WEBVISU : direct IEC variable] ADM100W L1 Max Load *)
  WEBVISU_OUTPUT_L1_L2_VOLTAGE_PHASE_ANGLE : DUT_Union_Real_Word;  (* [WEBVISU : direct IEC variable] ADM100W L1-L2 Voltage Phase Angle | deg *)
  WEBVISU_OUTPUT_L2_L3_VOLTAGE : DUT_Union_Real_Word;  (* [WEBVISU : direct IEC variable] ADM100W L2-L3 Voltage | V *)
  WEBVISU_OUTPUT_L2_N_VOLTAGE : DUT_Union_Real_Word;  (* [WEBVISU : direct IEC variable] ADM100W L2-N Voltage | V *)
  WEBVISU_OUTPUT_L2_CURRENT : DUT_Union_Real_Word;  (* [WEBVISU : direct IEC variable] ADM100W L2 Current | A *)
  WEBVISU_OUTPUT_L2_ACTIVE_POWER : DUT_Union_Real_Word;  (* [WEBVISU : direct IEC variable] ADM100W L2 Active Power *)
  WEBVISU_OUTPUT_L2_APPARENT_POWER : DUT_Union_Real_Word;  (* [WEBVISU : direct IEC variable] ADM100W L2 Apparent Power *)
  WEBVISU_OUTPUT_L2_REACTIVE_POWER : DUT_Union_Real_Word;  (* [WEBVISU : direct IEC variable] ADM100W L2 Reactive Power *)
  WEBVISU_OUTPUT_L2_CURRENT_PHASE_ANGLE : DUT_Union_Real_Word;  (* [WEBVISU : direct IEC variable] ADM100W L2 Current Phase Angle | deg *)
  WEBVISU_OUTPUT_L2_POWER_FACTOR : DUT_Union_Real_Word;  (* [WEBVISU : direct IEC variable] ADM100W L2 Power Factor *)
  WEBVISU_OUTPUT_L2_VOLTAGE_THD : DUT_Union_Real_Word;  (* [WEBVISU : direct IEC variable] ADM100W L2 Voltage THD | % *)
  WEBVISU_OUTPUT_L2_CURRENT_THD : DUT_Union_Real_Word;  (* [WEBVISU : direct IEC variable] ADM100W L2 Current THD | % *)
  WEBVISU_OUTPUT_L2_MAX_LOAD : DUT_Union_Real_Word;  (* [WEBVISU : direct IEC variable] ADM100W L2 Max Load *)
  WEBVISU_OUTPUT_L1_L3_VOLTAGE_PHASE_ANGLE : DUT_Union_Real_Word;  (* [WEBVISU : direct IEC variable] ADM100W L1-L3 Voltage Phase Angle | deg *)
  WEBVISU_OUTPUT_L3_L1_VOLTAGE : DUT_Union_Real_Word;  (* [WEBVISU : direct IEC variable] ADM100W L3-L1 Voltage | V *)
  WEBVISU_OUTPUT_L3_N_VOLTAGE : DUT_Union_Real_Word;  (* [WEBVISU : direct IEC variable] ADM100W L3-N Voltage | V *)
  WEBVISU_OUTPUT_L3_CURRENT : DUT_Union_Real_Word;  (* [WEBVISU : direct IEC variable] ADM100W L3 Current | A *)
  WEBVISU_OUTPUT_L3_ACTIVE_POWER : DUT_Union_Real_Word;  (* [WEBVISU : direct IEC variable] ADM100W L3 Active Power *)
  WEBVISU_OUTPUT_L3_APPARENT_POWER : DUT_Union_Real_Word;  (* [WEBVISU : direct IEC variable] ADM100W L3 Apparent Power *)
  WEBVISU_OUTPUT_L3_REACTIVE_POWER : DUT_Union_Real_Word;  (* [WEBVISU : direct IEC variable] ADM100W L3 Reactive Power *)
  WEBVISU_OUTPUT_L3_CURRENT_PHASE_ANGLE : DUT_Union_Real_Word;  (* [WEBVISU : direct IEC variable] ADM100W L3 Current Phase Angle | deg *)
  WEBVISU_OUTPUT_L3_POWER_FACTOR : DUT_Union_Real_Word;  (* [WEBVISU : direct IEC variable] ADM100W L3 Power Factor *)
  WEBVISU_OUTPUT_L3_VOLTAGE_THD : DUT_Union_Real_Word;  (* [WEBVISU : direct IEC variable] ADM100W L3 Voltage THD | % *)
  WEBVISU_OUTPUT_L3_CURRENT_THD : DUT_Union_Real_Word;  (* [WEBVISU : direct IEC variable] ADM100W L3 Current THD | % *)
  WEBVISU_OUTPUT_L3_MAX_LOAD : DUT_Union_Real_Word;  (* [WEBVISU : direct IEC variable] ADM100W L3 Max Load *)
  WEBVISU_OUTPUT_INTERNAL_TEMPERATURE : DUT_Union_Real_Word;  (* [WEBVISU : direct IEC variable] ADM100W Internal Temperature *)
  WEBVISU_OUTPUT_ACTIVE_ENERGY : DUT_Union_Real_Word;  (* [WEBVISU : direct IEC variable] ADM100W Active Energy *)
  WEBVISU_OUTPUT_APPARENT_ENERGY : DUT_Union_Real_Word;  (* [WEBVISU : direct IEC variable] ADM100W Apparent Energy *)
  WEBVISU_OUTPUT_REACTIVE_ENERGY : DUT_Union_Real_Word;  (* [WEBVISU : direct IEC variable] ADM100W Reactive Energy *)
  WEBVISU_OUTPUT_TOTAL_ACTIVE_POWER : DUT_Union_Real_Word;  (* [WEBVISU : direct IEC variable] ADM100W Total Active Power *)
  WEBVISU_OUTPUT_TOTAL_APPARENT_POWER : DUT_Union_Real_Word;  (* [WEBVISU : direct IEC variable] ADM100W Total Apparent Power *)
  WEBVISU_OUTPUT_TOTAL_REACTIVE_POWER : DUT_Union_Real_Word;  (* [WEBVISU : direct IEC variable] ADM100W Total Reactive Power *)
  WEBVISU_OUTPUT_ALL_PHASE_POWER_FACTOR : DUT_Union_Real_Word;  (* [WEBVISU : direct IEC variable] ADM100W All Phase Power Factor *)
  WEBVISU_OUTPUT_LOCAL_FUXA_ACTIVE : BOOL;  (* Effective FUXA local mode (masked by WEBVISU and HMI priority) *)
  WEBVISU_OUTPUT_LOCAL_HMI_ACTIVE : BOOL;  (* Effective HMI local mode (masked by WEBVISU priority) *)
END_STRUCT;
END_TYPE

TYPE DUT_EXC_ADM100W : STRUCT
  EXC_OUTPUT_FREQUENCY : REAL;  (* [EXC : to other equipment] Hz *)
  EXC_OUTPUT_L1_N_VOLTAGE : REAL;  (* V *)
  EXC_OUTPUT_L1_CURRENT : REAL;  (* A *)
  EXC_OUTPUT_L1_ACTIVE_POWER : REAL;  (* W *)
  EXC_OUTPUT_L1_APPARENT_POWER : REAL;  (* VA *)
  EXC_OUTPUT_L1_REACTIVE_POWER : REAL;  (* VAr *)
  EXC_OUTPUT_L1_POWER_FACTOR : REAL;  (* - *)
  EXC_OUTPUT_L1_VOLTAGE_THD : REAL;  (* % *)
  EXC_OUTPUT_L1_CURRENT_THD : REAL;  (* % *)
  EXC_OUTPUT_L1_MAX_LOAD : REAL;  (* % of 60 A *)
  EXC_OUTPUT_INTERNAL_TEMPERATURE : REAL;  (* degC *)
  EXC_OUTPUT_ACTIVE_ENERGY : REAL;  (* kWh *)
  EXC_OUTPUT_DATA_VALID : BOOL;  (* FALSE = values not usable. Not managed yet (no Modbus diagnostic) *)
  UPI_INPUT_GLOBAL_LOCAL_FUXA : BOOL;  (* [UPI : functional units to equipment] From UPI_LOCAL_FUXA : global FUXA local active *)
  UPI_INPUT_GLOBAL_LOCAL_HMI : BOOL;  (* From UPI_LOCAL_HMI : global HMI local active *)
  UPI_INPUT_GLOBAL_LOCAL_WEBVISU : BOOL;  (* From UPI_LOCAL_WEBVISU : global WEBVISU local active *)
END_STRUCT;
END_TYPE

TYPE DUT_COM_DIP1500 : STRUCT
  COM_INPUT_IR : ARRAY[0..4] OF WORD;  (* [COM : Modbus RTU, input (equipment to PLC)] Input registers 0x3001..0x3005 *)
  COM_INPUT_HR_COUNTERS : ARRAY[0..3] OF WORD;  (* Holding registers 0x4007..0x400A (read) *)
  COM_OUTPUT_COILS : ARRAY[0..3] OF BOOL;  (* [COM : Modbus RTU, output (PLC to equipment)] Coils 0x0001..0x0004 *)
  COM_OUTPUT_HR_CMD : ARRAY[0..5] OF WORD;  (* Holding registers 0x4001..0x4006 (write) *)
  COM_OUTPUT_HR_CONFIG : ARRAY[0..6] OF WORD;  (* Holding registers 0x400B..0x4011 (write) *)
  COM_OUTPUT_CMD_TRIGGER : BOOL;  (* Rising edge trigger of the command write channel(s), mapped in the Modbus slave I/O mapping *)
  COM_OUTPUT_CONFIG_TRIGGER : BOOL;  (* Rising edge trigger of the configuration write channel, mapped in the Modbus slave I/O mapping *)
  SCADA_INPUT_MOTOR_START_STOP : BOOL;  (* [SCADA (FUXA) : input (to PLC)] Coil 3 | DIP1500 Motor Start Stop *)
  SCADA_INPUT_MOTOR_DIRECTION : BOOL;  (* Coil 4 | DIP1500 Motor Direction *)
  SCADA_INPUT_FLASH_SAVE : BOOL;  (* Coil 5 | DIP1500 Flash Save *)
  SCADA_INPUT_OPERATION_MODE : BOOL;  (* Coil 6 | DIP1500 Operation Mode *)
  SCADA_INPUT_PARAM_WRITE_ENABLE : BOOL;  (* Coil 7 | DIP1500 Parameter Write Enable *)
  SCADA_INPUT_LOCAL_REQUEST : BOOL;  (* Coil 10 | DIP1500 Local Request *)
  SCADA_INPUT_AUTO_REQUEST : BOOL;  (* Coil 11 | DIP1500 Auto Request *)
  SCADA_INPUT_FOOT_SWITCH_INPUT_MODE : WORD;  (* HR 9 | DIP1500 Foot Switch Input Mode *)
  SCADA_INPUT_LIQUID_LEVEL_INPUT_MODE : WORD;  (* HR 10 | DIP1500 Liquid Level Input Mode *)
  SCADA_INPUT_STATE_OUTPUT_MODE : WORD;  (* HR 11 | DIP1500 State Output Mode *)
  SCADA_INPUT_COMMUNICATION_ADDRESS : WORD;  (* HR 12 | DIP1500 Communication Address *)
  SCADA_INPUT_BAUD_RATE_INDEX : WORD;  (* HR 13 | DIP1500 Baud Rate Index | index *)
  SCADA_INPUT_MOTOR_SPEED : DUT_Union_Real_Word;  (* HR 1-2 | DIP1500 Motor Speed | rpm *)
  SCADA_INPUT_MAX_MOTOR_SPEED : DUT_Union_Real_Word;  (* HR 3-4 | DIP1500 Max Motor Speed | rpm *)
  SCADA_INPUT_RUN_TIME_OR_VOLUME_SETPOINT : DUT_Union_Real_Word;  (* HR 5-6 | DIP1500 Run Time Or Volume Setpoint | ms (time mode) / ml (volume mode) *)
  SCADA_INPUT_FLOW_RATE_OR_SPEED_CALIBRATION_COEFFICIENT : DUT_Union_Real_Word;  (* HR 7-8 | DIP1500 Flow Rate Or Speed Calibration Coefficient | ml/min or rpm *)
  SCADA_OUTPUT_LOCAL_FUXA_ACTIVE : BOOL;  (* [SCADA (FUXA) : output (from PLC)] DI 10015 | DIP1500 Local FUXA Active *)
  SCADA_OUTPUT_LOCAL_HMI_ACTIVE : BOOL;  (* DI 10016 | DIP1500 Local HMI Active *)
  SCADA_OUTPUT_FIRMWARE_VERSION : WORD;  (* IR 91 | DIP1500 Firmware Version | 3+5+8 bits (major+minor+revision) *)
  SCADA_OUTPUT_HARDWARE_VERSION : WORD;  (* IR 92 | DIP1500 Hardware Version | 3+5+8 bits (major+minor+revision) *)
  SCADA_OUTPUT_TEMPERATURE : WORD;  (* IR 93 | DIP1500 Temperature | degC | (raw - 500) / 10 *)
  SCADA_OUTPUT_FLOAT_LEVEL_ALARM : WORD;  (* IR 94 | DIP1500 Float Level Alarm *)
  SCADA_OUTPUT_DIGITAL_OUTPUT_VALUE : WORD;  (* IR 95 | DIP1500 Digital Output Value *)
  SCADA_OUTPUT_REAL_TIME_RUN_TIME_OR_VOLUME : DUT_Union_Real_Word;  (* IR 96-97 | DIP1500 Real-Time Run Time Or Volume | ms (time mode) / ml (volume mode) *)
  SCADA_OUTPUT_ACCUMULATED_RUN_TIME_OR_VOLUME : DUT_Union_Real_Word;  (* IR 98-99 | DIP1500 Accumulated Run Time Or Volume | ms (time mode) / ml (volume mode) *)
  HMI_INPUT_MOTOR_START_STOP : BOOL;  (* [HMI (local panel, FUXA address + 1000) : input (to PLC)] Coil 1003 | DIP1500 Motor Start Stop *)
  HMI_INPUT_MOTOR_DIRECTION : BOOL;  (* Coil 1004 | DIP1500 Motor Direction *)
  HMI_INPUT_FLASH_SAVE : BOOL;  (* Coil 1005 | DIP1500 Flash Save *)
  HMI_INPUT_OPERATION_MODE : BOOL;  (* Coil 1006 | DIP1500 Operation Mode *)
  HMI_INPUT_PARAM_WRITE_ENABLE : BOOL;  (* Coil 1007 | DIP1500 Parameter Write Enable *)
  HMI_INPUT_LOCAL_REQUEST : BOOL;  (* Coil 1010 | DIP1500 Local Request *)
  HMI_INPUT_AUTO_REQUEST : BOOL;  (* Coil 1011 | DIP1500 Auto Request *)
  HMI_INPUT_FOOT_SWITCH_INPUT_MODE : WORD;  (* HR 1009 | DIP1500 Foot Switch Input Mode *)
  HMI_INPUT_LIQUID_LEVEL_INPUT_MODE : WORD;  (* HR 1010 | DIP1500 Liquid Level Input Mode *)
  HMI_INPUT_STATE_OUTPUT_MODE : WORD;  (* HR 1011 | DIP1500 State Output Mode *)
  HMI_INPUT_COMMUNICATION_ADDRESS : WORD;  (* HR 1012 | DIP1500 Communication Address *)
  HMI_INPUT_BAUD_RATE_INDEX : WORD;  (* HR 1013 | DIP1500 Baud Rate Index | index *)
  HMI_INPUT_MOTOR_SPEED : DUT_Union_Real_Word;  (* HR 1001-1002 | DIP1500 Motor Speed | rpm *)
  HMI_INPUT_MAX_MOTOR_SPEED : DUT_Union_Real_Word;  (* HR 1003-1004 | DIP1500 Max Motor Speed | rpm *)
  HMI_INPUT_RUN_TIME_OR_VOLUME_SETPOINT : DUT_Union_Real_Word;  (* HR 1005-1006 | DIP1500 Run Time Or Volume Setpoint | ms (time mode) / ml (volume mode) *)
  HMI_INPUT_FLOW_RATE_OR_SPEED_CALIBRATION_COEFFICIENT : DUT_Union_Real_Word;  (* HR 1007-1008 | DIP1500 Flow Rate Or Speed Calibration Coefficient | ml/min or rpm *)
  HMI_OUTPUT_LOCAL_ACTIVE : BOOL;  (* [HMI (local panel, FUXA address + 1000) : output (from PLC)] DI 11016 | DIP1500 Local Active *)
  HMI_OUTPUT_FIRMWARE_VERSION : WORD;  (* IR 1091 | DIP1500 Firmware Version | 3+5+8 bits (major+minor+revision) *)
  HMI_OUTPUT_HARDWARE_VERSION : WORD;  (* IR 1092 | DIP1500 Hardware Version | 3+5+8 bits (major+minor+revision) *)
  HMI_OUTPUT_TEMPERATURE : WORD;  (* IR 1093 | DIP1500 Temperature | degC | (raw - 500) / 10 *)
  HMI_OUTPUT_FLOAT_LEVEL_ALARM : WORD;  (* IR 1094 | DIP1500 Float Level Alarm *)
  HMI_OUTPUT_DIGITAL_OUTPUT_VALUE : WORD;  (* IR 1095 | DIP1500 Digital Output Value *)
  HMI_OUTPUT_REAL_TIME_RUN_TIME_OR_VOLUME : DUT_Union_Real_Word;  (* IR 1096-1097 | DIP1500 Real-Time Run Time Or Volume | ms (time mode) / ml (volume mode) *)
  HMI_OUTPUT_ACCUMULATED_RUN_TIME_OR_VOLUME : DUT_Union_Real_Word;  (* IR 1098-1099 | DIP1500 Accumulated Run Time Or Volume | ms (time mode) / ml (volume mode) *)
  WEBVISU_INPUT_MOTOR_START_STOP : BOOL;  (* [WEBVISU : direct IEC variable] DIP1500 Motor Start Stop *)
  WEBVISU_INPUT_MOTOR_DIRECTION : BOOL;  (* [WEBVISU : direct IEC variable] DIP1500 Motor Direction *)
  WEBVISU_INPUT_FLASH_SAVE : BOOL;  (* [WEBVISU : direct IEC variable] DIP1500 Flash Save *)
  WEBVISU_INPUT_OPERATION_MODE : BOOL;  (* [WEBVISU : direct IEC variable] DIP1500 Operation Mode *)
  WEBVISU_INPUT_PARAM_WRITE_ENABLE : BOOL;  (* [WEBVISU : direct IEC variable] DIP1500 Parameter Write Enable *)
  WEBVISU_INPUT_LOCAL_REQUEST : BOOL;  (* [WEBVISU : direct IEC variable] DIP1500 Local Request *)
  WEBVISU_INPUT_AUTO_REQUEST : BOOL;  (* [WEBVISU : direct IEC variable] DIP1500 Auto Request *)
  WEBVISU_INPUT_FOOT_SWITCH_INPUT_MODE : WORD;  (* [WEBVISU : direct IEC variable] DIP1500 Foot Switch Input Mode *)
  WEBVISU_INPUT_LIQUID_LEVEL_INPUT_MODE : WORD;  (* [WEBVISU : direct IEC variable] DIP1500 Liquid Level Input Mode *)
  WEBVISU_INPUT_STATE_OUTPUT_MODE : WORD;  (* [WEBVISU : direct IEC variable] DIP1500 State Output Mode *)
  WEBVISU_INPUT_COMMUNICATION_ADDRESS : WORD;  (* [WEBVISU : direct IEC variable] DIP1500 Communication Address *)
  WEBVISU_INPUT_BAUD_RATE_INDEX : WORD;  (* [WEBVISU : direct IEC variable] DIP1500 Baud Rate Index | index *)
  WEBVISU_INPUT_MOTOR_SPEED : DUT_Union_Real_Word;  (* [WEBVISU : direct IEC variable] DIP1500 Motor Speed | rpm *)
  WEBVISU_INPUT_MAX_MOTOR_SPEED : DUT_Union_Real_Word;  (* [WEBVISU : direct IEC variable] DIP1500 Max Motor Speed | rpm *)
  WEBVISU_INPUT_RUN_TIME_OR_VOLUME_SETPOINT : DUT_Union_Real_Word;  (* [WEBVISU : direct IEC variable] DIP1500 Run Time Or Volume Setpoint | ms (time mode) / ml (volume mode) *)
  WEBVISU_INPUT_FLOW_RATE_OR_SPEED_CALIBRATION_COEFFICIENT : DUT_Union_Real_Word;  (* [WEBVISU : direct IEC variable] DIP1500 Flow Rate Or Speed Calibration Coefficient | ml/min or rpm *)
  WEBVISU_OUTPUT_LOCAL_ACTIVE : BOOL;  (* [WEBVISU : direct IEC variable] DIP1500 Local Active *)
  WEBVISU_OUTPUT_FIRMWARE_VERSION : WORD;  (* [WEBVISU : direct IEC variable] DIP1500 Firmware Version | 3+5+8 bits (major+minor+revision) *)
  WEBVISU_OUTPUT_HARDWARE_VERSION : WORD;  (* [WEBVISU : direct IEC variable] DIP1500 Hardware Version | 3+5+8 bits (major+minor+revision) *)
  WEBVISU_OUTPUT_TEMPERATURE : WORD;  (* [WEBVISU : direct IEC variable] DIP1500 Temperature | degC | (raw - 500) / 10 *)
  WEBVISU_OUTPUT_FLOAT_LEVEL_ALARM : WORD;  (* [WEBVISU : direct IEC variable] DIP1500 Float Level Alarm *)
  WEBVISU_OUTPUT_DIGITAL_OUTPUT_VALUE : WORD;  (* [WEBVISU : direct IEC variable] DIP1500 Digital Output Value *)
  WEBVISU_OUTPUT_REAL_TIME_RUN_TIME_OR_VOLUME : DUT_Union_Real_Word;  (* [WEBVISU : direct IEC variable] DIP1500 Real-Time Run Time Or Volume | ms (time mode) / ml (volume mode) *)
  WEBVISU_OUTPUT_ACCUMULATED_RUN_TIME_OR_VOLUME : DUT_Union_Real_Word;  (* [WEBVISU : direct IEC variable] DIP1500 Accumulated Run Time Or Volume | ms (time mode) / ml (volume mode) *)
  WEBVISU_OUTPUT_LOCAL_FUXA_ACTIVE : BOOL;  (* Effective FUXA local mode (masked by WEBVISU and HMI priority) *)
  WEBVISU_OUTPUT_LOCAL_HMI_ACTIVE : BOOL;  (* Effective HMI local mode (masked by WEBVISU priority) *)
END_STRUCT;
END_TYPE

TYPE DUT_EXC_DIP1500 : STRUCT
  UPI_INPUT_GLOBAL_LOCAL_FUXA : BOOL;  (* [UPI : functional units to equipment] From UPI_LOCAL_FUXA : global FUXA local active *)
  UPI_INPUT_GLOBAL_LOCAL_HMI : BOOL;  (* From UPI_LOCAL_HMI : global HMI local active *)
  UPI_INPUT_RUN : BOOL;  (* [UPI : commands used in auto mode] Auto mode command : run *)
  UPI_INPUT_CLOCKWISE : BOOL;  (* Auto mode command : 1 clockwise *)
  UPI_INPUT_VOLUME_MODE : BOOL;  (* Auto mode command : 0 time mode, 1 volume mode *)
  UPI_INPUT_SPEED : REAL;  (* Auto mode command : speed, rpm *)
  UPI_INPUT_RUN_SETPOINT : REAL;  (* Auto mode command : ms (time mode) or ml (volume mode), 0 = continuous *)
  UPI_INPUT_GLOBAL_LOCAL_WEBVISU : BOOL;  (* From UPI_LOCAL_WEBVISU : global WEBVISU local active *)
END_STRUCT;
END_TYPE

TYPE DUT_IO_DIP1500 : STRUCT
  SPARE : BOOL;  (* Placeholder, structure not used yet *)
END_STRUCT;
END_TYPE

TYPE DUT_PA_ADM100W : STRUCT
  SPARE : BOOL;  (* Placeholder, structure not used yet *)
END_STRUCT;
END_TYPE

TYPE DUT_PA_DOSENSOR : STRUCT
  SPARE : BOOL;  (* Placeholder, structure not used yet *)
END_STRUCT;
END_TYPE

TYPE DUT_PA_DIP1500 : STRUCT
  MAX_MOTOR_SPEED : REAL := 350;  (* [Pump configuration, default value = declaration value, kept in GVL_PA (persistent)] rpm. Max motor speed (pump register 0x4003) *)
  CALIBRATION_COEFFICIENT : REAL := 100;  (* ml/min or rpm. Flow / speed calibration coefficient (0x400B) *)
  FOOT_SWITCH_INPUT_MODE : WORD := 0;  (* Foot switch input mode (0x400D) *)
  LIQUID_LEVEL_INPUT_MODE : WORD := 100;  (* Liquid level input mode (0x400E) *)
  STATE_OUTPUT_MODE : WORD := 7;  (* State output mode (0x400F) *)
  COMMUNICATION_ADDRESS : WORD := 11;  (* Pump Modbus address, 1..31 (0x4010) *)
  BAUD_RATE_INDEX : WORD := 3;  (* 0=1200 .. 3=9600 .. 7=115200 (0x4011) *)
END_STRUCT;
END_TYPE

TYPE DUT_COM_UPI_LOCAL_HMI : STRUCT
  SCADA_OUTPUT_LOCAL_ACTIVE : BOOL;  (* [SCADA (FUXA) : output (from PLC)] DI 10020 | Global Local HMI Active *)
  HMI_INPUT_LOCAL_REQUEST : BOOL;  (* [HMI (local panel, FUXA address + 1000) : input (to PLC)] Coil 1014 | Global Local HMI Request *)
  HMI_INPUT_AUTO_REQUEST : BOOL;  (* Coil 1015 | Global Auto HMI Request *)
  HMI_OUTPUT_LOCAL_ACTIVE : BOOL;  (* [HMI (local panel, FUXA address + 1000) : output (from PLC)] DI 11020 | Global Local HMI Active *)
END_STRUCT;
END_TYPE

TYPE DUT_EXC_UPI_LOCAL_FUXA : STRUCT
  UPI_OUTPUT_LOCAL_ACTIVE : BOOL;  (* [UPI : to equipment] Global FUXA local active *)
END_STRUCT;
END_TYPE

TYPE DUT_EXC_UPI_LOCAL_HMI : STRUCT
  UPI_OUTPUT_LOCAL_ACTIVE : BOOL;  (* [UPI : to equipment] Global HMI local active *)
END_STRUCT;
END_TYPE

TYPE DUT_INT_UPI_LOCAL_FUXA : STRUCT
  LOCAL_REQUEST : BOOL;  (* Local request (pulse or maintained) *)
  AUTO_REQUEST : BOOL;  (* Auto request, releases the global local *)
  LOCAL_ACTIVE : BOOL;  (* Memory : global local active *)
END_STRUCT;
END_TYPE

TYPE DUT_INT_UPI_LOCAL_HMI : STRUCT
  LOCAL_REQUEST : BOOL;  (* Local request (pulse or maintained) *)
  AUTO_REQUEST : BOOL;  (* Auto request, releases the global local *)
  LOCAL_ACTIVE : BOOL;  (* Memory : global local active *)
END_STRUCT;
END_TYPE

TYPE DUT_COM_UPI_LOCAL_WEBVISU : STRUCT
  WEBVISU_INPUT_LOCAL_REQUEST : BOOL;  (* [WEBVISU (direct IEC variables) : input (to PLC)] Global Local WEBVISU Request *)
  WEBVISU_INPUT_AUTO_REQUEST : BOOL;  (* Global Auto WEBVISU Request *)
  WEBVISU_OUTPUT_LOCAL_ACTIVE : BOOL;  (* [WEBVISU (direct IEC variables) : output (from PLC)] Global Local WEBVISU Active *)
END_STRUCT;
END_TYPE

TYPE DUT_EXC_UPI_LOCAL_WEBVISU : STRUCT
  UPI_OUTPUT_LOCAL_ACTIVE : BOOL;  (* [UPI : to equipment] Global WEBVISU local active *)
END_STRUCT;
END_TYPE

TYPE DUT_INT_UPI_LOCAL_WEBVISU : STRUCT
  LOCAL_REQUEST : BOOL;  (* Local request (pulse or maintained) *)
  AUTO_REQUEST : BOOL;  (* Auto request, releases the global local *)
  LOCAL_ACTIVE : BOOL;  (* Memory : global local active *)
END_STRUCT;
END_TYPE

TYPE DUT_Union_Real_Word : UNION
  Real_value : REAL;
  Word_value : ARRAY[0..1] OF WORD;
END_UNION;
END_TYPE

FUNCTION_BLOCK FB_INST_ADM100W
  VAR_IN_OUT
    PA : DUT_PA_ADM100W;  (* Parameters (persistent, GVL_PA) *)
    COM : DUT_COM_ADM100W;  (* Communication : Modbus RTU (COM_), SCADA FUXA (SCADA_), HMI (HMI_) *)
    EXC : DUT_EXC_ADM100W;  (* Exchanges : other equipment (EXC_), functional units (UPI_) *)
    IO : DUT_IO_ADM100W;  (* Wired PLC I/O *)
  END_VAR
  VAR
    INTERN : DUT_INT_ADM100W;  (* Internal variables *)
  END_VAR

                  
//==============================================================================
// FB_INST_ADM100W
// Trumeter ADM100W power meter, Modbus RTU, 32-bit float MSW first (ABCD). No command : local mode is only reported
// 1. INPUTS     : requests, control mode, command source, equipment feedback -> INTERN
// 2. PROCESSING : on INTERN only
// 3. OUTPUTS    : INTERN -> COM / IO / EXC
// Control mode  : local WEBVISU > local HMI > local FUXA > auto (functional units)
//==============================================================================

//------------------------------------------------------------------------------
// 1. INPUTS
//------------------------------------------------------------------------------
	//--- Control mode requests (WEBVISU, HMI, FUXA, global UPI)
	INTERN.FUXA_LOCAL_REQUEST := COM.SCADA_INPUT_LOCAL_REQUEST;
	INTERN.FUXA_AUTO_REQUEST  := COM.SCADA_INPUT_AUTO_REQUEST;
	INTERN.HMI_LOCAL_REQUEST  := COM.HMI_INPUT_LOCAL_REQUEST;
	INTERN.HMI_AUTO_REQUEST   := COM.HMI_INPUT_AUTO_REQUEST;
	INTERN.GLOBAL_LOCAL_FUXA  := EXC.UPI_INPUT_GLOBAL_LOCAL_FUXA;
	INTERN.GLOBAL_LOCAL_HMI   := EXC.UPI_INPUT_GLOBAL_LOCAL_HMI;
	INTERN.WEBVISU_LOCAL_REQUEST := COM.WEBVISU_INPUT_LOCAL_REQUEST;
	INTERN.WEBVISU_AUTO_REQUEST  := COM.WEBVISU_INPUT_AUTO_REQUEST;
	INTERN.GLOBAL_LOCAL_WEBVISU  := EXC.UPI_INPUT_GLOBAL_LOCAL_WEBVISU;

	//--- Control mode
	// Individual memories : set by the local request, reset by the auto request (auto wins if both)
	IF INTERN.WEBVISU_LOCAL_REQUEST THEN
		INTERN.LOCAL_WEBVISU_INDIVIDUAL := TRUE;
	END_IF
	IF INTERN.WEBVISU_AUTO_REQUEST THEN
		INTERN.LOCAL_WEBVISU_INDIVIDUAL := FALSE;
	END_IF
	IF INTERN.HMI_LOCAL_REQUEST THEN
		INTERN.LOCAL_HMI_INDIVIDUAL := TRUE;
	END_IF
	IF INTERN.HMI_AUTO_REQUEST THEN
		INTERN.LOCAL_HMI_INDIVIDUAL := FALSE;
	END_IF
	IF INTERN.FUXA_LOCAL_REQUEST THEN
		INTERN.LOCAL_FUXA_INDIVIDUAL := TRUE;
	END_IF
	IF INTERN.FUXA_AUTO_REQUEST THEN
		INTERN.LOCAL_FUXA_INDIVIDUAL := FALSE;
	END_IF

	// Resulting mode : individual OR global, WEBVISU > HMI > FUXA > auto
	INTERN.LOCAL_WEBVISU := INTERN.LOCAL_WEBVISU_INDIVIDUAL OR INTERN.GLOBAL_LOCAL_WEBVISU;
	INTERN.LOCAL_HMI     := (INTERN.LOCAL_HMI_INDIVIDUAL OR INTERN.GLOBAL_LOCAL_HMI) AND NOT INTERN.LOCAL_WEBVISU;
	INTERN.LOCAL_FUXA    := (INTERN.LOCAL_FUXA_INDIVIDUAL OR INTERN.GLOBAL_LOCAL_FUXA) AND NOT INTERN.LOCAL_WEBVISU AND NOT INTERN.LOCAL_HMI;
	INTERN.AUTO          := NOT INTERN.LOCAL_WEBVISU AND NOT INTERN.LOCAL_HMI AND NOT INTERN.LOCAL_FUXA;

	//--- COM : alarms (coils 0..9)
	INTERN.ALARM_1  := COM.COM_INPUT_COILS[0].0;
	INTERN.ALARM_2  := COM.COM_INPUT_COILS[0].1;
	INTERN.ALARM_3  := COM.COM_INPUT_COILS[0].2;
	INTERN.ALARM_4  := COM.COM_INPUT_COILS[0].3;
	INTERN.ALARM_5  := COM.COM_INPUT_COILS[0].4;
	INTERN.ALARM_6  := COM.COM_INPUT_COILS[0].5;
	INTERN.ALARM_7  := COM.COM_INPUT_COILS[0].6;
	INTERN.ALARM_8  := COM.COM_INPUT_COILS[0].7;
	INTERN.ALARM_9  := COM.COM_INPUT_COILS[1].0;
	INTERN.ALARM_10 := COM.COM_INPUT_COILS[1].1;

	//--- COM : measures (input registers, MSW first)
	INTERN.FREQUENCY                 := FNC_WORDS_TO_REAL(High_word := COM.COM_INPUT_IR[0], Low_word := COM.COM_INPUT_IR[1]);
	INTERN.L1_L2_VOLTAGE             := FNC_WORDS_TO_REAL(High_word := COM.COM_INPUT_IR[2], Low_word := COM.COM_INPUT_IR[3]);
	INTERN.L1_N_VOLTAGE              := FNC_WORDS_TO_REAL(High_word := COM.COM_INPUT_IR[4], Low_word := COM.COM_INPUT_IR[5]);
	INTERN.L1_CURRENT                := FNC_WORDS_TO_REAL(High_word := COM.COM_INPUT_IR[6], Low_word := COM.COM_INPUT_IR[7]);
	INTERN.L1_ACTIVE_POWER           := FNC_WORDS_TO_REAL(High_word := COM.COM_INPUT_IR[8], Low_word := COM.COM_INPUT_IR[9]);
	INTERN.L1_APPARENT_POWER         := FNC_WORDS_TO_REAL(High_word := COM.COM_INPUT_IR[10], Low_word := COM.COM_INPUT_IR[11]);
	INTERN.L1_REACTIVE_POWER         := FNC_WORDS_TO_REAL(High_word := COM.COM_INPUT_IR[12], Low_word := COM.COM_INPUT_IR[13]);
	INTERN.L1_CURRENT_PHASE_ANGLE    := FNC_WORDS_TO_REAL(High_word := COM.COM_INPUT_IR[14], Low_word := COM.COM_INPUT_IR[15]);
	INTERN.L1_POWER_FACTOR           := FNC_WORDS_TO_REAL(High_word := COM.COM_INPUT_IR[16], Low_word := COM.COM_INPUT_IR[17]);
	INTERN.L1_VOLTAGE_THD            := FNC_WORDS_TO_REAL(High_word := COM.COM_INPUT_IR[18], Low_word := COM.COM_INPUT_IR[19]);
	INTERN.L1_CURRENT_THD            := FNC_WORDS_TO_REAL(High_word := COM.COM_INPUT_IR[20], Low_word := COM.COM_INPUT_IR[21]);
	INTERN.L1_MAX_LOAD               := FNC_WORDS_TO_REAL(High_word := COM.COM_INPUT_IR[22], Low_word := COM.COM_INPUT_IR[23]);
	INTERN.L1_L2_VOLTAGE_PHASE_ANGLE := FNC_WORDS_TO_REAL(High_word := COM.COM_INPUT_IR[24], Low_word := COM.COM_INPUT_IR[25]);
	INTERN.L2_L3_VOLTAGE             := FNC_WORDS_TO_REAL(High_word := COM.COM_INPUT_IR[26], Low_word := COM.COM_INPUT_IR[27]);
	INTERN.L2_N_VOLTAGE              := FNC_WORDS_TO_REAL(High_word := COM.COM_INPUT_IR[28], Low_word := COM.COM_INPUT_IR[29]);
	INTERN.L2_CURRENT                := FNC_WORDS_TO_REAL(High_word := COM.COM_INPUT_IR[30], Low_word := COM.COM_INPUT_IR[31]);
	INTERN.L2_ACTIVE_POWER           := FNC_WORDS_TO_REAL(High_word := COM.COM_INPUT_IR[32], Low_word := COM.COM_INPUT_IR[33]);
	INTERN.L2_APPARENT_POWER         := FNC_WORDS_TO_REAL(High_word := COM.COM_INPUT_IR[34], Low_word := COM.COM_INPUT_IR[35]);
	INTERN.L2_REACTIVE_POWER         := FNC_WORDS_TO_REAL(High_word := COM.COM_INPUT_IR[36], Low_word := COM.COM_INPUT_IR[37]);
	INTERN.L2_CURRENT_PHASE_ANGLE    := FNC_WORDS_TO_REAL(High_word := COM.COM_INPUT_IR[38], Low_word := COM.COM_INPUT_IR[39]);
	INTERN.L2_POWER_FACTOR           := FNC_WORDS_TO_REAL(High_word := COM.COM_INPUT_IR[40], Low_word := COM.COM_INPUT_IR[41]);
	INTERN.L2_VOLTAGE_THD            := FNC_WORDS_TO_REAL(High_word := COM.COM_INPUT_IR[42], Low_word := COM.COM_INPUT_IR[43]);
	INTERN.L2_CURRENT_THD            := FNC_WORDS_TO_REAL(High_word := COM.COM_INPUT_IR[44], Low_word := COM.COM_INPUT_IR[45]);
	INTERN.L2_MAX_LOAD               := FNC_WORDS_TO_REAL(High_word := COM.COM_INPUT_IR[46], Low_word := COM.COM_INPUT_IR[47]);
	INTERN.L1_L3_VOLTAGE_PHASE_ANGLE := FNC_WORDS_TO_REAL(High_word := COM.COM_INPUT_IR[48], Low_word := COM.COM_INPUT_IR[49]);
	INTERN.L3_L1_VOLTAGE             := FNC_WORDS_TO_REAL(High_word := COM.COM_INPUT_IR[50], Low_word := COM.COM_INPUT_IR[51]);
	INTERN.L3_N_VOLTAGE              := FNC_WORDS_TO_REAL(High_word := COM.COM_INPUT_IR[52], Low_word := COM.COM_INPUT_IR[53]);
	INTERN.L3_CURRENT                := FNC_WORDS_TO_REAL(High_word := COM.COM_INPUT_IR[54], Low_word := COM.COM_INPUT_IR[55]);
	INTERN.L3_ACTIVE_POWER           := FNC_WORDS_TO_REAL(High_word := COM.COM_INPUT_IR[56], Low_word := COM.COM_INPUT_IR[57]);
	INTERN.L3_APPARENT_POWER         := FNC_WORDS_TO_REAL(High_word := COM.COM_INPUT_IR[58], Low_word := COM.COM_INPUT_IR[59]);
	INTERN.L3_REACTIVE_POWER         := FNC_WORDS_TO_REAL(High_word := COM.COM_INPUT_IR[60], Low_word := COM.COM_INPUT_IR[61]);
	INTERN.L3_CURRENT_PHASE_ANGLE    := FNC_WORDS_TO_REAL(High_word := COM.COM_INPUT_IR[62], Low_word := COM.COM_INPUT_IR[63]);
	INTERN.L3_POWER_FACTOR           := FNC_WORDS_TO_REAL(High_word := COM.COM_INPUT_IR[64], Low_word := COM.COM_INPUT_IR[65]);
	INTERN.L3_VOLTAGE_THD            := FNC_WORDS_TO_REAL(High_word := COM.COM_INPUT_IR[66], Low_word := COM.COM_INPUT_IR[67]);
	INTERN.L3_CURRENT_THD            := FNC_WORDS_TO_REAL(High_word := COM.COM_INPUT_IR[68], Low_word := COM.COM_INPUT_IR[69]);
	INTERN.L3_MAX_LOAD               := FNC_WORDS_TO_REAL(High_word := COM.COM_INPUT_IR[70], Low_word := COM.COM_INPUT_IR[71]);
	INTERN.INTERNAL_TEMPERATURE      := FNC_WORDS_TO_REAL(High_word := COM.COM_INPUT_IR[72], Low_word := COM.COM_INPUT_IR[73]);
	INTERN.ACTIVE_ENERGY             := FNC_WORDS_TO_REAL(High_word := COM.COM_INPUT_IR[74], Low_word := COM.COM_INPUT_IR[75]);
	INTERN.APPARENT_ENERGY           := FNC_WORDS_TO_REAL(High_word := COM.COM_INPUT_IR[76], Low_word := COM.COM_INPUT_IR[77]);
	INTERN.REACTIVE_ENERGY           := FNC_WORDS_TO_REAL(High_word := COM.COM_INPUT_IR[78], Low_word := COM.COM_INPUT_IR[79]);
	INTERN.TOTAL_ACTIVE_POWER        := FNC_WORDS_TO_REAL(High_word := COM.COM_INPUT_IR[80], Low_word := COM.COM_INPUT_IR[81]);
	INTERN.TOTAL_APPARENT_POWER      := FNC_WORDS_TO_REAL(High_word := COM.COM_INPUT_IR[82], Low_word := COM.COM_INPUT_IR[83]);
	INTERN.TOTAL_REACTIVE_POWER      := FNC_WORDS_TO_REAL(High_word := COM.COM_INPUT_IR[84], Low_word := COM.COM_INPUT_IR[85]);
	INTERN.ALL_PHASE_POWER_FACTOR    := FNC_WORDS_TO_REAL(High_word := COM.COM_INPUT_IR[86], Low_word := COM.COM_INPUT_IR[87]);


//------------------------------------------------------------------------------
// 2. PROCESSING
//------------------------------------------------------------------------------
	// Nothing


//------------------------------------------------------------------------------
// 3. OUTPUTS
//------------------------------------------------------------------------------
	//--- COM : control mode status to SCADA, HMI and WEBVISU
	COM.SCADA_OUTPUT_LOCAL_FUXA_ACTIVE := INTERN.LOCAL_FUXA;
	COM.SCADA_OUTPUT_LOCAL_HMI_ACTIVE  := INTERN.LOCAL_HMI;
	COM.HMI_OUTPUT_LOCAL_ACTIVE        := INTERN.LOCAL_HMI;
	COM.WEBVISU_OUTPUT_LOCAL_ACTIVE        := INTERN.LOCAL_WEBVISU;
	COM.WEBVISU_OUTPUT_LOCAL_HMI_ACTIVE  := INTERN.LOCAL_HMI;
	COM.WEBVISU_OUTPUT_LOCAL_FUXA_ACTIVE := INTERN.LOCAL_FUXA;

	//--- EXC
	EXC.EXC_OUTPUT_FREQUENCY            := INTERN.FREQUENCY;
	EXC.EXC_OUTPUT_L1_N_VOLTAGE         := INTERN.L1_N_VOLTAGE;
	EXC.EXC_OUTPUT_L1_CURRENT           := INTERN.L1_CURRENT;
	EXC.EXC_OUTPUT_L1_ACTIVE_POWER      := INTERN.L1_ACTIVE_POWER;
	EXC.EXC_OUTPUT_L1_APPARENT_POWER    := INTERN.L1_APPARENT_POWER;
	EXC.EXC_OUTPUT_L1_REACTIVE_POWER    := INTERN.L1_REACTIVE_POWER;
	EXC.EXC_OUTPUT_L1_POWER_FACTOR      := INTERN.L1_POWER_FACTOR;
	EXC.EXC_OUTPUT_L1_VOLTAGE_THD       := INTERN.L1_VOLTAGE_THD;
	EXC.EXC_OUTPUT_L1_CURRENT_THD       := INTERN.L1_CURRENT_THD;
	EXC.EXC_OUTPUT_L1_MAX_LOAD          := INTERN.L1_MAX_LOAD;
	EXC.EXC_OUTPUT_INTERNAL_TEMPERATURE := INTERN.INTERNAL_TEMPERATURE;
	EXC.EXC_OUTPUT_ACTIVE_ENERGY        := INTERN.ACTIVE_ENERGY;
	// EXC.EXC_OUTPUT_DATA_VALID : not managed yet (no Modbus diagnostic)

	//--- COM : alarms to SCADA, HMI and WEBVISU
	COM.SCADA_OUTPUT_ALARM_1_STATUS  := INTERN.ALARM_1;
	COM.HMI_OUTPUT_ALARM_1_STATUS    := INTERN.ALARM_1;
	COM.WEBVISU_OUTPUT_ALARM_1_STATUS    := INTERN.ALARM_1;
	COM.SCADA_OUTPUT_ALARM_2_STATUS  := INTERN.ALARM_2;
	COM.HMI_OUTPUT_ALARM_2_STATUS    := INTERN.ALARM_2;
	COM.WEBVISU_OUTPUT_ALARM_2_STATUS    := INTERN.ALARM_2;
	COM.SCADA_OUTPUT_ALARM_3_STATUS  := INTERN.ALARM_3;
	COM.HMI_OUTPUT_ALARM_3_STATUS    := INTERN.ALARM_3;
	COM.WEBVISU_OUTPUT_ALARM_3_STATUS    := INTERN.ALARM_3;
	COM.SCADA_OUTPUT_ALARM_4_STATUS  := INTERN.ALARM_4;
	COM.HMI_OUTPUT_ALARM_4_STATUS    := INTERN.ALARM_4;
	COM.WEBVISU_OUTPUT_ALARM_4_STATUS    := INTERN.ALARM_4;
	COM.SCADA_OUTPUT_ALARM_5_STATUS  := INTERN.ALARM_5;
	COM.HMI_OUTPUT_ALARM_5_STATUS    := INTERN.ALARM_5;
	COM.WEBVISU_OUTPUT_ALARM_5_STATUS    := INTERN.ALARM_5;
	COM.SCADA_OUTPUT_ALARM_6_STATUS  := INTERN.ALARM_6;
	COM.HMI_OUTPUT_ALARM_6_STATUS    := INTERN.ALARM_6;
	COM.WEBVISU_OUTPUT_ALARM_6_STATUS    := INTERN.ALARM_6;
	COM.SCADA_OUTPUT_ALARM_7_STATUS  := INTERN.ALARM_7;
	COM.HMI_OUTPUT_ALARM_7_STATUS    := INTERN.ALARM_7;
	COM.WEBVISU_OUTPUT_ALARM_7_STATUS    := INTERN.ALARM_7;
	COM.SCADA_OUTPUT_ALARM_8_STATUS  := INTERN.ALARM_8;
	COM.HMI_OUTPUT_ALARM_8_STATUS    := INTERN.ALARM_8;
	COM.WEBVISU_OUTPUT_ALARM_8_STATUS    := INTERN.ALARM_8;
	COM.SCADA_OUTPUT_ALARM_9_STATUS  := INTERN.ALARM_9;
	COM.HMI_OUTPUT_ALARM_9_STATUS    := INTERN.ALARM_9;
	COM.WEBVISU_OUTPUT_ALARM_9_STATUS    := INTERN.ALARM_9;
	COM.SCADA_OUTPUT_ALARM_10_STATUS := INTERN.ALARM_10;
	COM.HMI_OUTPUT_ALARM_10_STATUS   := INTERN.ALARM_10;
	COM.WEBVISU_OUTPUT_ALARM_10_STATUS   := INTERN.ALARM_10;

	//--- COM : measures to SCADA, HMI and WEBVISU
	COM.SCADA_OUTPUT_FREQUENCY.Real_value                 := INTERN.FREQUENCY;
	COM.HMI_OUTPUT_FREQUENCY.Real_value                   := INTERN.FREQUENCY;
	COM.WEBVISU_OUTPUT_FREQUENCY.Real_value                   := INTERN.FREQUENCY;
	COM.SCADA_OUTPUT_L1_L2_VOLTAGE.Real_value             := INTERN.L1_L2_VOLTAGE;
	COM.HMI_OUTPUT_L1_L2_VOLTAGE.Real_value               := INTERN.L1_L2_VOLTAGE;
	COM.WEBVISU_OUTPUT_L1_L2_VOLTAGE.Real_value               := INTERN.L1_L2_VOLTAGE;
	COM.SCADA_OUTPUT_L1_N_VOLTAGE.Real_value              := INTERN.L1_N_VOLTAGE;
	COM.HMI_OUTPUT_L1_N_VOLTAGE.Real_value                := INTERN.L1_N_VOLTAGE;
	COM.WEBVISU_OUTPUT_L1_N_VOLTAGE.Real_value                := INTERN.L1_N_VOLTAGE;
	COM.SCADA_OUTPUT_L1_CURRENT.Real_value                := INTERN.L1_CURRENT;
	COM.HMI_OUTPUT_L1_CURRENT.Real_value                  := INTERN.L1_CURRENT;
	COM.WEBVISU_OUTPUT_L1_CURRENT.Real_value                  := INTERN.L1_CURRENT;
	COM.SCADA_OUTPUT_L1_ACTIVE_POWER.Real_value           := INTERN.L1_ACTIVE_POWER;
	COM.HMI_OUTPUT_L1_ACTIVE_POWER.Real_value             := INTERN.L1_ACTIVE_POWER;
	COM.WEBVISU_OUTPUT_L1_ACTIVE_POWER.Real_value             := INTERN.L1_ACTIVE_POWER;
	COM.SCADA_OUTPUT_L1_APPARENT_POWER.Real_value         := INTERN.L1_APPARENT_POWER;
	COM.HMI_OUTPUT_L1_APPARENT_POWER.Real_value           := INTERN.L1_APPARENT_POWER;
	COM.WEBVISU_OUTPUT_L1_APPARENT_POWER.Real_value           := INTERN.L1_APPARENT_POWER;
	COM.SCADA_OUTPUT_L1_REACTIVE_POWER.Real_value         := INTERN.L1_REACTIVE_POWER;
	COM.HMI_OUTPUT_L1_REACTIVE_POWER.Real_value           := INTERN.L1_REACTIVE_POWER;
	COM.WEBVISU_OUTPUT_L1_REACTIVE_POWER.Real_value           := INTERN.L1_REACTIVE_POWER;
	COM.SCADA_OUTPUT_L1_CURRENT_PHASE_ANGLE.Real_value    := INTERN.L1_CURRENT_PHASE_ANGLE;
	COM.HMI_OUTPUT_L1_CURRENT_PHASE_ANGLE.Real_value      := INTERN.L1_CURRENT_PHASE_ANGLE;
	COM.WEBVISU_OUTPUT_L1_CURRENT_PHASE_ANGLE.Real_value      := INTERN.L1_CURRENT_PHASE_ANGLE;
	COM.SCADA_OUTPUT_L1_POWER_FACTOR.Real_value           := INTERN.L1_POWER_FACTOR;
	COM.HMI_OUTPUT_L1_POWER_FACTOR.Real_value             := INTERN.L1_POWER_FACTOR;
	COM.WEBVISU_OUTPUT_L1_POWER_FACTOR.Real_value             := INTERN.L1_POWER_FACTOR;
	COM.SCADA_OUTPUT_L1_VOLTAGE_THD.Real_value            := INTERN.L1_VOLTAGE_THD;
	COM.HMI_OUTPUT_L1_VOLTAGE_THD.Real_value              := INTERN.L1_VOLTAGE_THD;
	COM.WEBVISU_OUTPUT_L1_VOLTAGE_THD.Real_value              := INTERN.L1_VOLTAGE_THD;
	COM.SCADA_OUTPUT_L1_CURRENT_THD.Real_value            := INTERN.L1_CURRENT_THD;
	COM.HMI_OUTPUT_L1_CURRENT_THD.Real_value              := INTERN.L1_CURRENT_THD;
	COM.WEBVISU_OUTPUT_L1_CURRENT_THD.Real_value              := INTERN.L1_CURRENT_THD;
	COM.SCADA_OUTPUT_L1_MAX_LOAD.Real_value               := INTERN.L1_MAX_LOAD;
	COM.HMI_OUTPUT_L1_MAX_LOAD.Real_value                 := INTERN.L1_MAX_LOAD;
	COM.WEBVISU_OUTPUT_L1_MAX_LOAD.Real_value                 := INTERN.L1_MAX_LOAD;
	COM.SCADA_OUTPUT_L1_L2_VOLTAGE_PHASE_ANGLE.Real_value := INTERN.L1_L2_VOLTAGE_PHASE_ANGLE;
	COM.HMI_OUTPUT_L1_L2_VOLTAGE_PHASE_ANGLE.Real_value   := INTERN.L1_L2_VOLTAGE_PHASE_ANGLE;
	COM.WEBVISU_OUTPUT_L1_L2_VOLTAGE_PHASE_ANGLE.Real_value   := INTERN.L1_L2_VOLTAGE_PHASE_ANGLE;
	COM.SCADA_OUTPUT_L2_L3_VOLTAGE.Real_value             := INTERN.L2_L3_VOLTAGE;
	COM.HMI_OUTPUT_L2_L3_VOLTAGE.Real_value               := INTERN.L2_L3_VOLTAGE;
	COM.WEBVISU_OUTPUT_L2_L3_VOLTAGE.Real_value               := INTERN.L2_L3_VOLTAGE;
	COM.SCADA_OUTPUT_L2_N_VOLTAGE.Real_value              := INTERN.L2_N_VOLTAGE;
	COM.HMI_OUTPUT_L2_N_VOLTAGE.Real_value                := INTERN.L2_N_VOLTAGE;
	COM.WEBVISU_OUTPUT_L2_N_VOLTAGE.Real_value                := INTERN.L2_N_VOLTAGE;
	COM.SCADA_OUTPUT_L2_CURRENT.Real_value                := INTERN.L2_CURRENT;
	COM.HMI_OUTPUT_L2_CURRENT.Real_value                  := INTERN.L2_CURRENT;
	COM.WEBVISU_OUTPUT_L2_CURRENT.Real_value                  := INTERN.L2_CURRENT;
	COM.SCADA_OUTPUT_L2_ACTIVE_POWER.Real_value           := INTERN.L2_ACTIVE_POWER;
	COM.HMI_OUTPUT_L2_ACTIVE_POWER.Real_value             := INTERN.L2_ACTIVE_POWER;
	COM.WEBVISU_OUTPUT_L2_ACTIVE_POWER.Real_value             := INTERN.L2_ACTIVE_POWER;
	COM.SCADA_OUTPUT_L2_APPARENT_POWER.Real_value         := INTERN.L2_APPARENT_POWER;
	COM.HMI_OUTPUT_L2_APPARENT_POWER.Real_value           := INTERN.L2_APPARENT_POWER;
	COM.WEBVISU_OUTPUT_L2_APPARENT_POWER.Real_value           := INTERN.L2_APPARENT_POWER;
	COM.SCADA_OUTPUT_L2_REACTIVE_POWER.Real_value         := INTERN.L2_REACTIVE_POWER;
	COM.HMI_OUTPUT_L2_REACTIVE_POWER.Real_value           := INTERN.L2_REACTIVE_POWER;
	COM.WEBVISU_OUTPUT_L2_REACTIVE_POWER.Real_value           := INTERN.L2_REACTIVE_POWER;
	COM.SCADA_OUTPUT_L2_CURRENT_PHASE_ANGLE.Real_value    := INTERN.L2_CURRENT_PHASE_ANGLE;
	COM.HMI_OUTPUT_L2_CURRENT_PHASE_ANGLE.Real_value      := INTERN.L2_CURRENT_PHASE_ANGLE;
	COM.WEBVISU_OUTPUT_L2_CURRENT_PHASE_ANGLE.Real_value      := INTERN.L2_CURRENT_PHASE_ANGLE;
	COM.SCADA_OUTPUT_L2_POWER_FACTOR.Real_value           := INTERN.L2_POWER_FACTOR;
	COM.HMI_OUTPUT_L2_POWER_FACTOR.Real_value             := INTERN.L2_POWER_FACTOR;
	COM.WEBVISU_OUTPUT_L2_POWER_FACTOR.Real_value             := INTERN.L2_POWER_FACTOR;
	COM.SCADA_OUTPUT_L2_VOLTAGE_THD.Real_value            := INTERN.L2_VOLTAGE_THD;
	COM.HMI_OUTPUT_L2_VOLTAGE_THD.Real_value              := INTERN.L2_VOLTAGE_THD;
	COM.WEBVISU_OUTPUT_L2_VOLTAGE_THD.Real_value              := INTERN.L2_VOLTAGE_THD;
	COM.SCADA_OUTPUT_L2_CURRENT_THD.Real_value            := INTERN.L2_CURRENT_THD;
	COM.HMI_OUTPUT_L2_CURRENT_THD.Real_value              := INTERN.L2_CURRENT_THD;
	COM.WEBVISU_OUTPUT_L2_CURRENT_THD.Real_value              := INTERN.L2_CURRENT_THD;
	COM.SCADA_OUTPUT_L2_MAX_LOAD.Real_value               := INTERN.L2_MAX_LOAD;
	COM.HMI_OUTPUT_L2_MAX_LOAD.Real_value                 := INTERN.L2_MAX_LOAD;
	COM.WEBVISU_OUTPUT_L2_MAX_LOAD.Real_value                 := INTERN.L2_MAX_LOAD;
	COM.SCADA_OUTPUT_L1_L3_VOLTAGE_PHASE_ANGLE.Real_value := INTERN.L1_L3_VOLTAGE_PHASE_ANGLE;
	COM.HMI_OUTPUT_L1_L3_VOLTAGE_PHASE_ANGLE.Real_value   := INTERN.L1_L3_VOLTAGE_PHASE_ANGLE;
	COM.WEBVISU_OUTPUT_L1_L3_VOLTAGE_PHASE_ANGLE.Real_value   := INTERN.L1_L3_VOLTAGE_PHASE_ANGLE;
	COM.SCADA_OUTPUT_L3_L1_VOLTAGE.Real_value             := INTERN.L3_L1_VOLTAGE;
	COM.HMI_OUTPUT_L3_L1_VOLTAGE.Real_value               := INTERN.L3_L1_VOLTAGE;
	COM.WEBVISU_OUTPUT_L3_L1_VOLTAGE.Real_value               := INTERN.L3_L1_VOLTAGE;
	COM.SCADA_OUTPUT_L3_N_VOLTAGE.Real_value              := INTERN.L3_N_VOLTAGE;
	COM.HMI_OUTPUT_L3_N_VOLTAGE.Real_value                := INTERN.L3_N_VOLTAGE;
	COM.WEBVISU_OUTPUT_L3_N_VOLTAGE.Real_value                := INTERN.L3_N_VOLTAGE;
	COM.SCADA_OUTPUT_L3_CURRENT.Real_value                := INTERN.L3_CURRENT;
	COM.HMI_OUTPUT_L3_CURRENT.Real_value                  := INTERN.L3_CURRENT;
	COM.WEBVISU_OUTPUT_L3_CURRENT.Real_value                  := INTERN.L3_CURRENT;
	COM.SCADA_OUTPUT_L3_ACTIVE_POWER.Real_value           := INTERN.L3_ACTIVE_POWER;
	COM.HMI_OUTPUT_L3_ACTIVE_POWER.Real_value             := INTERN.L3_ACTIVE_POWER;
	COM.WEBVISU_OUTPUT_L3_ACTIVE_POWER.Real_value             := INTERN.L3_ACTIVE_POWER;
	COM.SCADA_OUTPUT_L3_APPARENT_POWER.Real_value         := INTERN.L3_APPARENT_POWER;
	COM.HMI_OUTPUT_L3_APPARENT_POWER.Real_value           := INTERN.L3_APPARENT_POWER;
	COM.WEBVISU_OUTPUT_L3_APPARENT_POWER.Real_value           := INTERN.L3_APPARENT_POWER;
	COM.SCADA_OUTPUT_L3_REACTIVE_POWER.Real_value         := INTERN.L3_REACTIVE_POWER;
	COM.HMI_OUTPUT_L3_REACTIVE_POWER.Real_value           := INTERN.L3_REACTIVE_POWER;
	COM.WEBVISU_OUTPUT_L3_REACTIVE_POWER.Real_value           := INTERN.L3_REACTIVE_POWER;
	COM.SCADA_OUTPUT_L3_CURRENT_PHASE_ANGLE.Real_value    := INTERN.L3_CURRENT_PHASE_ANGLE;
	COM.HMI_OUTPUT_L3_CURRENT_PHASE_ANGLE.Real_value      := INTERN.L3_CURRENT_PHASE_ANGLE;
	COM.WEBVISU_OUTPUT_L3_CURRENT_PHASE_ANGLE.Real_value      := INTERN.L3_CURRENT_PHASE_ANGLE;
	COM.SCADA_OUTPUT_L3_POWER_FACTOR.Real_value           := INTERN.L3_POWER_FACTOR;
	COM.HMI_OUTPUT_L3_POWER_FACTOR.Real_value             := INTERN.L3_POWER_FACTOR;
	COM.WEBVISU_OUTPUT_L3_POWER_FACTOR.Real_value             := INTERN.L3_POWER_FACTOR;
	COM.SCADA_OUTPUT_L3_VOLTAGE_THD.Real_value            := INTERN.L3_VOLTAGE_THD;
	COM.HMI_OUTPUT_L3_VOLTAGE_THD.Real_value              := INTERN.L3_VOLTAGE_THD;
	COM.WEBVISU_OUTPUT_L3_VOLTAGE_THD.Real_value              := INTERN.L3_VOLTAGE_THD;
	COM.SCADA_OUTPUT_L3_CURRENT_THD.Real_value            := INTERN.L3_CURRENT_THD;
	COM.HMI_OUTPUT_L3_CURRENT_THD.Real_value              := INTERN.L3_CURRENT_THD;
	COM.WEBVISU_OUTPUT_L3_CURRENT_THD.Real_value              := INTERN.L3_CURRENT_THD;
	COM.SCADA_OUTPUT_L3_MAX_LOAD.Real_value               := INTERN.L3_MAX_LOAD;
	COM.HMI_OUTPUT_L3_MAX_LOAD.Real_value                 := INTERN.L3_MAX_LOAD;
	COM.WEBVISU_OUTPUT_L3_MAX_LOAD.Real_value                 := INTERN.L3_MAX_LOAD;
	COM.SCADA_OUTPUT_INTERNAL_TEMPERATURE.Real_value      := INTERN.INTERNAL_TEMPERATURE;
	COM.HMI_OUTPUT_INTERNAL_TEMPERATURE.Real_value        := INTERN.INTERNAL_TEMPERATURE;
	COM.WEBVISU_OUTPUT_INTERNAL_TEMPERATURE.Real_value        := INTERN.INTERNAL_TEMPERATURE;
	COM.SCADA_OUTPUT_ACTIVE_ENERGY.Real_value             := INTERN.ACTIVE_ENERGY;
	COM.HMI_OUTPUT_ACTIVE_ENERGY.Real_value               := INTERN.ACTIVE_ENERGY;
	COM.WEBVISU_OUTPUT_ACTIVE_ENERGY.Real_value               := INTERN.ACTIVE_ENERGY;
	COM.SCADA_OUTPUT_APPARENT_ENERGY.Real_value           := INTERN.APPARENT_ENERGY;
	COM.HMI_OUTPUT_APPARENT_ENERGY.Real_value             := INTERN.APPARENT_ENERGY;
	COM.WEBVISU_OUTPUT_APPARENT_ENERGY.Real_value             := INTERN.APPARENT_ENERGY;
	COM.SCADA_OUTPUT_REACTIVE_ENERGY.Real_value           := INTERN.REACTIVE_ENERGY;
	COM.HMI_OUTPUT_REACTIVE_ENERGY.Real_value             := INTERN.REACTIVE_ENERGY;
	COM.WEBVISU_OUTPUT_REACTIVE_ENERGY.Real_value             := INTERN.REACTIVE_ENERGY;
	COM.SCADA_OUTPUT_TOTAL_ACTIVE_POWER.Real_value        := INTERN.TOTAL_ACTIVE_POWER;
	COM.HMI_OUTPUT_TOTAL_ACTIVE_POWER.Real_value          := INTERN.TOTAL_ACTIVE_POWER;
	COM.WEBVISU_OUTPUT_TOTAL_ACTIVE_POWER.Real_value          := INTERN.TOTAL_ACTIVE_POWER;
	COM.SCADA_OUTPUT_TOTAL_APPARENT_POWER.Real_value      := INTERN.TOTAL_APPARENT_POWER;
	COM.HMI_OUTPUT_TOTAL_APPARENT_POWER.Real_value        := INTERN.TOTAL_APPARENT_POWER;
	COM.WEBVISU_OUTPUT_TOTAL_APPARENT_POWER.Real_value        := INTERN.TOTAL_APPARENT_POWER;
	COM.SCADA_OUTPUT_TOTAL_REACTIVE_POWER.Real_value      := INTERN.TOTAL_REACTIVE_POWER;
	COM.HMI_OUTPUT_TOTAL_REACTIVE_POWER.Real_value        := INTERN.TOTAL_REACTIVE_POWER;
	COM.WEBVISU_OUTPUT_TOTAL_REACTIVE_POWER.Real_value        := INTERN.TOTAL_REACTIVE_POWER;
	COM.SCADA_OUTPUT_ALL_PHASE_POWER_FACTOR.Real_value    := INTERN.ALL_PHASE_POWER_FACTOR;
	COM.HMI_OUTPUT_ALL_PHASE_POWER_FACTOR.Real_value      := INTERN.ALL_PHASE_POWER_FACTOR;
	COM.WEBVISU_OUTPUT_ALL_PHASE_POWER_FACTOR.Real_value      := INTERN.ALL_PHASE_POWER_FACTOR;


                
END_FUNCTION_BLOCK

FUNCTION_BLOCK FB_INST_DOSENSOR
  VAR_IN_OUT
    PA : DUT_PA_DOSENSOR;  (* Parameters (persistent, GVL_PA) *)
    COM : DUT_COM_DOSENSOR;  (* Communication : Modbus RTU (COM_), SCADA FUXA (SCADA_), HMI (HMI_) *)
    EXC : DUT_EXC_DOSENSOR;  (* Exchanges : other equipment (EXC_), functional units (UPI_) *)
    IO : DUT_IO_DOSENSOR;  (* Wired PLC I/O *)
  END_VAR
  VAR
    INTERN : DUT_INT_DOSENSOR;  (* Internal variables *)
    TP_CALIB_HIGH : TP;  (* High calibration pulse *)
    TP_CALIB_LOW : TP;  (* Low calibration pulse *)
    TP_CALIB_DONE : TP;  (* Calibration done message *)
  END_VAR

                  
//==============================================================================
// FB_INST_DOSENSOR
// Dissolved oxygen sensor, analog signal + fault input + 2 calibration outputs
// 1. INPUTS     : requests, control mode, command source, equipment feedback -> INTERN
// 2. PROCESSING : on INTERN only
// 3. OUTPUTS    : INTERN -> COM / IO / EXC
// Control mode  : local WEBVISU > local HMI > local FUXA > auto (functional units)
//==============================================================================

//------------------------------------------------------------------------------
// 1. INPUTS
//------------------------------------------------------------------------------
	//--- Control mode requests (WEBVISU, HMI, FUXA, global UPI)
	INTERN.FUXA_LOCAL_REQUEST := COM.SCADA_INPUT_LOCAL_REQUEST;
	INTERN.FUXA_AUTO_REQUEST  := COM.SCADA_INPUT_AUTO_REQUEST;
	INTERN.HMI_LOCAL_REQUEST  := COM.HMI_INPUT_LOCAL_REQUEST;
	INTERN.HMI_AUTO_REQUEST   := COM.HMI_INPUT_AUTO_REQUEST;
	INTERN.GLOBAL_LOCAL_FUXA  := EXC.UPI_INPUT_GLOBAL_LOCAL_FUXA;
	INTERN.GLOBAL_LOCAL_HMI   := EXC.UPI_INPUT_GLOBAL_LOCAL_HMI;
	INTERN.WEBVISU_LOCAL_REQUEST := COM.WEBVISU_INPUT_LOCAL_REQUEST;
	INTERN.WEBVISU_AUTO_REQUEST  := COM.WEBVISU_INPUT_AUTO_REQUEST;
	INTERN.GLOBAL_LOCAL_WEBVISU  := EXC.UPI_INPUT_GLOBAL_LOCAL_WEBVISU;
	//--- Control mode
	// Individual memories : set by the local request, reset by the auto request (auto wins if both)
	IF INTERN.WEBVISU_LOCAL_REQUEST THEN
		INTERN.LOCAL_WEBVISU_INDIVIDUAL := TRUE;
	END_IF
	IF INTERN.WEBVISU_AUTO_REQUEST THEN
		INTERN.LOCAL_WEBVISU_INDIVIDUAL := FALSE;
	END_IF
	IF INTERN.HMI_LOCAL_REQUEST THEN
		INTERN.LOCAL_HMI_INDIVIDUAL := TRUE;
	END_IF
	IF INTERN.HMI_AUTO_REQUEST THEN
		INTERN.LOCAL_HMI_INDIVIDUAL := FALSE;
	END_IF
	IF INTERN.FUXA_LOCAL_REQUEST THEN
		INTERN.LOCAL_FUXA_INDIVIDUAL := TRUE;
	END_IF
	IF INTERN.FUXA_AUTO_REQUEST THEN
		INTERN.LOCAL_FUXA_INDIVIDUAL := FALSE;
	END_IF

	// Resulting mode : individual OR global, WEBVISU > HMI > FUXA > auto
	INTERN.LOCAL_WEBVISU := INTERN.LOCAL_WEBVISU_INDIVIDUAL OR INTERN.GLOBAL_LOCAL_WEBVISU;
	INTERN.LOCAL_HMI     := (INTERN.LOCAL_HMI_INDIVIDUAL OR INTERN.GLOBAL_LOCAL_HMI) AND NOT INTERN.LOCAL_WEBVISU;
	INTERN.LOCAL_FUXA    := (INTERN.LOCAL_FUXA_INDIVIDUAL OR INTERN.GLOBAL_LOCAL_FUXA) AND NOT INTERN.LOCAL_WEBVISU AND NOT INTERN.LOCAL_HMI;
	INTERN.AUTO          := NOT INTERN.LOCAL_WEBVISU AND NOT INTERN.LOCAL_HMI AND NOT INTERN.LOCAL_FUXA;

	//--- Command source : calibration requests
	IF INTERN.LOCAL_WEBVISU THEN
		INTERN.CALIB_HIGH_REQUEST := COM.WEBVISU_INPUT_CALIBRATION_HIGH;
		INTERN.CALIB_LOW_REQUEST  := COM.WEBVISU_INPUT_CALIBRATION_LOW;
	ELSIF INTERN.LOCAL_HMI THEN
		INTERN.CALIB_HIGH_REQUEST := COM.HMI_INPUT_CALIBRATION_HIGH;
		INTERN.CALIB_LOW_REQUEST  := COM.HMI_INPUT_CALIBRATION_LOW;
	ELSIF INTERN.LOCAL_FUXA THEN
		INTERN.CALIB_HIGH_REQUEST := COM.SCADA_INPUT_CALIBRATION_HIGH;
		INTERN.CALIB_LOW_REQUEST  := COM.SCADA_INPUT_CALIBRATION_LOW;
	ELSE
		// Auto : functional units (UPI)
		INTERN.CALIB_HIGH_REQUEST := FALSE;
		INTERN.CALIB_LOW_REQUEST  := FALSE;
	END_IF

	//--- IO
	INTERN.SIGNAL_RAW := IO.INPUT_SIGNAL;
	INTERN.FAULT      := IO.INPUT_SENSOR_FAULT;


//------------------------------------------------------------------------------
// 2. PROCESSING
//------------------------------------------------------------------------------
	//--- Signal scaling
	INTERN.SIGNAL := (DWORD_TO_REAL(INTERN.SIGNAL_RAW * 40) / 65535) - 8;

	//--- Calibration : 1 s pulse to the sensor, 5 s "done" message
	TP_CALIB_HIGH(IN := INTERN.CALIB_HIGH_REQUEST, PT := T#1S);
	TP_CALIB_LOW(IN := INTERN.CALIB_LOW_REQUEST, PT := T#1S);
	TP_CALIB_DONE(IN := TP_CALIB_HIGH.Q OR TP_CALIB_LOW.Q, PT := T#5S);

	INTERN.CALIB_HIGH := TP_CALIB_HIGH.Q;
	INTERN.CALIB_LOW  := TP_CALIB_LOW.Q;
	INTERN.CALIB_DONE := TP_CALIB_DONE.Q;


//------------------------------------------------------------------------------
// 3. OUTPUTS
//------------------------------------------------------------------------------
	//--- COM : control mode status to SCADA, HMI and WEBVISU
	COM.SCADA_OUTPUT_LOCAL_FUXA_ACTIVE := INTERN.LOCAL_FUXA;
	COM.SCADA_OUTPUT_LOCAL_HMI_ACTIVE  := INTERN.LOCAL_HMI;
	COM.HMI_OUTPUT_LOCAL_ACTIVE        := INTERN.LOCAL_HMI;
	COM.WEBVISU_OUTPUT_LOCAL_ACTIVE        := INTERN.LOCAL_WEBVISU;
	COM.WEBVISU_OUTPUT_LOCAL_HMI_ACTIVE  := INTERN.LOCAL_HMI;
	COM.WEBVISU_OUTPUT_LOCAL_FUXA_ACTIVE := INTERN.LOCAL_FUXA;

	//--- EXC
	EXC.EXC_OUTPUT_SIGNAL := INTERN.SIGNAL;

	//--- IO
	IO.OUTPUT_CALIBRATION_HIGH := INTERN.CALIB_HIGH;
	IO.OUTPUT_CALIBRATION_LOW  := INTERN.CALIB_LOW;

	//--- COM : feedback to SCADA, HMI and WEBVISU
	COM.SCADA_OUTPUT_SIGNAL.Real_value := INTERN.SIGNAL;
	COM.HMI_OUTPUT_SIGNAL.Real_value   := INTERN.SIGNAL;
	COM.WEBVISU_OUTPUT_SIGNAL.Real_value   := INTERN.SIGNAL;
	COM.SCADA_OUTPUT_FAULT             := INTERN.FAULT;
	COM.HMI_OUTPUT_FAULT               := INTERN.FAULT;
	COM.WEBVISU_OUTPUT_FAULT               := INTERN.FAULT;
	COM.SCADA_OUTPUT_CALIBRATION_DONE  := INTERN.CALIB_DONE;
	COM.HMI_OUTPUT_CALIBRATION_DONE    := INTERN.CALIB_DONE;
	COM.WEBVISU_OUTPUT_CALIBRATION_DONE    := INTERN.CALIB_DONE;


                
END_FUNCTION_BLOCK

FUNCTION_BLOCK FB_INST_DIP1500
  VAR_IN_OUT
    PA : DUT_PA_DIP1500;  (* Parameters (persistent, GVL_PA) *)
    COM : DUT_COM_DIP1500;  (* Communication : Modbus RTU (COM_), SCADA FUXA (SCADA_), HMI (HMI_) *)
    EXC : DUT_EXC_DIP1500;  (* Exchanges : other equipment (EXC_), functional units (UPI_) *)
    IO : DUT_IO_DIP1500;  (* Wired PLC I/O *)
  END_VAR
  VAR
    INTERN : DUT_INT_DIP1500;  (* Internal variables *)
    TON_PULSE : TON;  (* Square wave timer *)
    TOF_CMD_WINDOW : TOF;  (* Command write window *)
    R_TRIG_FLASH : R_TRIG;  (* Flash save request edge *)
    TP_FLASH : TP;  (* Flash save pulse *)
  END_VAR

                  
//==============================================================================
// FB_INST_DIP1500
// Kamoer DIP1500 peristaltic pump, Modbus RTU, 32-bit low word first (CDAB)
// 1. INPUTS     : requests, control mode, command source, equipment feedback -> INTERN
// 2. PROCESSING : on INTERN only
// 3. OUTPUTS    : INTERN -> COM / IO / EXC
// Parameters    : pump configuration in PA (persistent), changed from the active local supervision
// Control mode  : local WEBVISU > local HMI > local FUXA > auto (functional units)
//==============================================================================

//------------------------------------------------------------------------------
// 1. INPUTS
//------------------------------------------------------------------------------
	//--- Control mode requests (WEBVISU, HMI, FUXA, global UPI)
	INTERN.FUXA_LOCAL_REQUEST := COM.SCADA_INPUT_LOCAL_REQUEST;
	INTERN.FUXA_AUTO_REQUEST  := COM.SCADA_INPUT_AUTO_REQUEST;
	INTERN.HMI_LOCAL_REQUEST  := COM.HMI_INPUT_LOCAL_REQUEST;
	INTERN.HMI_AUTO_REQUEST   := COM.HMI_INPUT_AUTO_REQUEST;
	INTERN.GLOBAL_LOCAL_FUXA  := EXC.UPI_INPUT_GLOBAL_LOCAL_FUXA;
	INTERN.GLOBAL_LOCAL_HMI   := EXC.UPI_INPUT_GLOBAL_LOCAL_HMI;
	INTERN.WEBVISU_LOCAL_REQUEST := COM.WEBVISU_INPUT_LOCAL_REQUEST;
	INTERN.WEBVISU_AUTO_REQUEST  := COM.WEBVISU_INPUT_AUTO_REQUEST;
	INTERN.GLOBAL_LOCAL_WEBVISU  := EXC.UPI_INPUT_GLOBAL_LOCAL_WEBVISU;

	//--- Control mode
	// Individual memories : set by the local request, reset by the auto request (auto wins if both)
	IF INTERN.WEBVISU_LOCAL_REQUEST THEN
		INTERN.LOCAL_WEBVISU_INDIVIDUAL := TRUE;
	END_IF
	IF INTERN.WEBVISU_AUTO_REQUEST THEN
		INTERN.LOCAL_WEBVISU_INDIVIDUAL := FALSE;
	END_IF
	IF INTERN.HMI_LOCAL_REQUEST THEN
		INTERN.LOCAL_HMI_INDIVIDUAL := TRUE;
	END_IF
	IF INTERN.HMI_AUTO_REQUEST THEN
		INTERN.LOCAL_HMI_INDIVIDUAL := FALSE;
	END_IF
	IF INTERN.FUXA_LOCAL_REQUEST THEN
		INTERN.LOCAL_FUXA_INDIVIDUAL := TRUE;
	END_IF
	IF INTERN.FUXA_AUTO_REQUEST THEN
		INTERN.LOCAL_FUXA_INDIVIDUAL := FALSE;
	END_IF

	// Resulting mode : individual OR global, WEBVISU > HMI > FUXA > auto
	INTERN.LOCAL_WEBVISU := INTERN.LOCAL_WEBVISU_INDIVIDUAL OR INTERN.GLOBAL_LOCAL_WEBVISU;
	INTERN.LOCAL_HMI     := (INTERN.LOCAL_HMI_INDIVIDUAL OR INTERN.GLOBAL_LOCAL_HMI) AND NOT INTERN.LOCAL_WEBVISU;
	INTERN.LOCAL_FUXA    := (INTERN.LOCAL_FUXA_INDIVIDUAL OR INTERN.GLOBAL_LOCAL_FUXA) AND NOT INTERN.LOCAL_WEBVISU AND NOT INTERN.LOCAL_HMI;
	INTERN.AUTO          := NOT INTERN.LOCAL_WEBVISU AND NOT INTERN.LOCAL_HMI AND NOT INTERN.LOCAL_FUXA;

	//--- Command source : local WEBVISU > local HMI > local FUXA > auto (UPI)
	IF INTERN.LOCAL_WEBVISU THEN
		INTERN.CMD_RUN            := COM.WEBVISU_INPUT_MOTOR_START_STOP;
		INTERN.CMD_CLOCKWISE      := COM.WEBVISU_INPUT_MOTOR_DIRECTION;
		INTERN.CMD_VOLUME_MODE    := COM.WEBVISU_INPUT_OPERATION_MODE;
		INTERN.CMD_SPEED          := COM.WEBVISU_INPUT_MOTOR_SPEED.Real_value;
		INTERN.CMD_RUN_SETPOINT   := COM.WEBVISU_INPUT_RUN_TIME_OR_VOLUME_SETPOINT.Real_value;
		INTERN.PARAM_WRITE_ENABLE := COM.WEBVISU_INPUT_PARAM_WRITE_ENABLE;
		INTERN.FLASH_SAVE_REQUEST := COM.WEBVISU_INPUT_FLASH_SAVE;
	ELSIF INTERN.LOCAL_HMI THEN
		INTERN.CMD_RUN            := COM.HMI_INPUT_MOTOR_START_STOP;
		INTERN.CMD_CLOCKWISE      := COM.HMI_INPUT_MOTOR_DIRECTION;
		INTERN.CMD_VOLUME_MODE    := COM.HMI_INPUT_OPERATION_MODE;
		INTERN.CMD_SPEED          := COM.HMI_INPUT_MOTOR_SPEED.Real_value;
		INTERN.CMD_RUN_SETPOINT   := COM.HMI_INPUT_RUN_TIME_OR_VOLUME_SETPOINT.Real_value;
		INTERN.PARAM_WRITE_ENABLE := COM.HMI_INPUT_PARAM_WRITE_ENABLE;
		INTERN.FLASH_SAVE_REQUEST := COM.HMI_INPUT_FLASH_SAVE;
	ELSIF INTERN.LOCAL_FUXA THEN
		INTERN.CMD_RUN            := COM.SCADA_INPUT_MOTOR_START_STOP;
		INTERN.CMD_CLOCKWISE      := COM.SCADA_INPUT_MOTOR_DIRECTION;
		INTERN.CMD_VOLUME_MODE    := COM.SCADA_INPUT_OPERATION_MODE;
		INTERN.CMD_SPEED          := COM.SCADA_INPUT_MOTOR_SPEED.Real_value;
		INTERN.CMD_RUN_SETPOINT   := COM.SCADA_INPUT_RUN_TIME_OR_VOLUME_SETPOINT.Real_value;
		INTERN.PARAM_WRITE_ENABLE := COM.SCADA_INPUT_PARAM_WRITE_ENABLE;
		INTERN.FLASH_SAVE_REQUEST := COM.SCADA_INPUT_FLASH_SAVE;
	ELSE
		// Auto : functional units (UPI)
		INTERN.CMD_RUN            := EXC.UPI_INPUT_RUN;
		INTERN.CMD_CLOCKWISE      := EXC.UPI_INPUT_CLOCKWISE;
		INTERN.CMD_VOLUME_MODE    := EXC.UPI_INPUT_VOLUME_MODE;
		INTERN.CMD_SPEED          := EXC.UPI_INPUT_SPEED;
		INTERN.CMD_RUN_SETPOINT   := EXC.UPI_INPUT_RUN_SETPOINT;
		INTERN.PARAM_WRITE_ENABLE := FALSE;                        // configuration is never written in auto
		INTERN.FLASH_SAVE_REQUEST := FALSE;
	END_IF

	//--- Parameter source : values typed in the active local supervision (nothing in auto)
	IF INTERN.LOCAL_WEBVISU THEN
		INTERN.SRC_MAX_MOTOR_SPEED         := COM.WEBVISU_INPUT_MAX_MOTOR_SPEED.Real_value;
		INTERN.SRC_CALIBRATION_COEFFICIENT := COM.WEBVISU_INPUT_FLOW_RATE_OR_SPEED_CALIBRATION_COEFFICIENT.Real_value;
		INTERN.SRC_FOOT_SWITCH_INPUT_MODE  := COM.WEBVISU_INPUT_FOOT_SWITCH_INPUT_MODE;
		INTERN.SRC_LIQUID_LEVEL_INPUT_MODE := COM.WEBVISU_INPUT_LIQUID_LEVEL_INPUT_MODE;
		INTERN.SRC_STATE_OUTPUT_MODE       := COM.WEBVISU_INPUT_STATE_OUTPUT_MODE;
		INTERN.SRC_COMMUNICATION_ADDRESS   := COM.WEBVISU_INPUT_COMMUNICATION_ADDRESS;
		INTERN.SRC_BAUD_RATE_INDEX         := COM.WEBVISU_INPUT_BAUD_RATE_INDEX;
	ELSIF INTERN.LOCAL_HMI THEN
		INTERN.SRC_MAX_MOTOR_SPEED         := COM.HMI_INPUT_MAX_MOTOR_SPEED.Real_value;
		INTERN.SRC_CALIBRATION_COEFFICIENT := COM.HMI_INPUT_FLOW_RATE_OR_SPEED_CALIBRATION_COEFFICIENT.Real_value;
		INTERN.SRC_FOOT_SWITCH_INPUT_MODE  := COM.HMI_INPUT_FOOT_SWITCH_INPUT_MODE;
		INTERN.SRC_LIQUID_LEVEL_INPUT_MODE := COM.HMI_INPUT_LIQUID_LEVEL_INPUT_MODE;
		INTERN.SRC_STATE_OUTPUT_MODE       := COM.HMI_INPUT_STATE_OUTPUT_MODE;
		INTERN.SRC_COMMUNICATION_ADDRESS   := COM.HMI_INPUT_COMMUNICATION_ADDRESS;
		INTERN.SRC_BAUD_RATE_INDEX         := COM.HMI_INPUT_BAUD_RATE_INDEX;
	ELSIF INTERN.LOCAL_FUXA THEN
		INTERN.SRC_MAX_MOTOR_SPEED         := COM.SCADA_INPUT_MAX_MOTOR_SPEED.Real_value;
		INTERN.SRC_CALIBRATION_COEFFICIENT := COM.SCADA_INPUT_FLOW_RATE_OR_SPEED_CALIBRATION_COEFFICIENT.Real_value;
		INTERN.SRC_FOOT_SWITCH_INPUT_MODE  := COM.SCADA_INPUT_FOOT_SWITCH_INPUT_MODE;
		INTERN.SRC_LIQUID_LEVEL_INPUT_MODE := COM.SCADA_INPUT_LIQUID_LEVEL_INPUT_MODE;
		INTERN.SRC_STATE_OUTPUT_MODE       := COM.SCADA_INPUT_STATE_OUTPUT_MODE;
		INTERN.SRC_COMMUNICATION_ADDRESS   := COM.SCADA_INPUT_COMMUNICATION_ADDRESS;
		INTERN.SRC_BAUD_RATE_INDEX         := COM.SCADA_INPUT_BAUD_RATE_INDEX;
	END_IF

	//--- COM : input registers 0x3001..0x3005
	INTERN.FBK_FIRMWARE_VERSION := COM.COM_INPUT_IR[0];
	INTERN.FBK_HARDWARE_VERSION := COM.COM_INPUT_IR[1];
	INTERN.FBK_TEMPERATURE      := COM.COM_INPUT_IR[2];
	INTERN.FBK_LEVEL_ALARM      := COM.COM_INPUT_IR[3];
	INTERN.FBK_DIGITAL_OUTPUT   := COM.COM_INPUT_IR[4];

	//--- COM : run counters 0x4007..0x400A (format depends on mode)
	IF INTERN.CMD_VOLUME_MODE THEN
		// Volume mode : 32-bit REAL (ml)
		INTERN.FBK_RUN_ACTUAL := FNC_WORDS_TO_REAL(High_word := COM.COM_INPUT_HR_COUNTERS[1], Low_word := COM.COM_INPUT_HR_COUNTERS[0]);
		INTERN.FBK_RUN_TOTAL  := FNC_WORDS_TO_REAL(High_word := COM.COM_INPUT_HR_COUNTERS[3], Low_word := COM.COM_INPUT_HR_COUNTERS[2]);
	ELSE
		// Time mode : 32-bit UDINT (ms)
		INTERN.UDINT_TEMP     := SHL(WORD_TO_UDINT(COM.COM_INPUT_HR_COUNTERS[1]), 16) OR WORD_TO_UDINT(COM.COM_INPUT_HR_COUNTERS[0]);
		INTERN.FBK_RUN_ACTUAL := UDINT_TO_REAL(INTERN.UDINT_TEMP);
		INTERN.UDINT_TEMP     := SHL(WORD_TO_UDINT(COM.COM_INPUT_HR_COUNTERS[3]), 16) OR WORD_TO_UDINT(COM.COM_INPUT_HR_COUNTERS[2]);
		INTERN.FBK_RUN_TOTAL  := UDINT_TO_REAL(INTERN.UDINT_TEMP);
	END_IF


//------------------------------------------------------------------------------
// 2. PROCESSING
//------------------------------------------------------------------------------
	//--- Parameters (PA) : a value changed in the active supervision is saved in PA
	// PA is persistent : it keeps its value after a restart or a download. Default = declaration value.
	// The cycle where the source changes is ignored, so switching mode never overwrites PA.
	INTERN.SOURCE_CHANGED := (INTERN.LOCAL_WEBVISU <> INTERN.PREV_LOCAL_WEBVISU)
	                         OR (INTERN.LOCAL_HMI <> INTERN.PREV_LOCAL_HMI)
	                         OR (INTERN.LOCAL_FUXA <> INTERN.PREV_LOCAL_FUXA);
	INTERN.PREV_LOCAL_WEBVISU := INTERN.LOCAL_WEBVISU;
	INTERN.PREV_LOCAL_HMI     := INTERN.LOCAL_HMI;
	INTERN.PREV_LOCAL_FUXA    := INTERN.LOCAL_FUXA;

	IF NOT INTERN.SOURCE_CHANGED THEN
		IF INTERN.SRC_MAX_MOTOR_SPEED <> INTERN.PREV_SRC_MAX_MOTOR_SPEED THEN
			PA.MAX_MOTOR_SPEED := INTERN.SRC_MAX_MOTOR_SPEED;
		END_IF
		IF INTERN.SRC_CALIBRATION_COEFFICIENT <> INTERN.PREV_SRC_CALIBRATION_COEFFICIENT THEN
			PA.CALIBRATION_COEFFICIENT := INTERN.SRC_CALIBRATION_COEFFICIENT;
		END_IF
		IF INTERN.SRC_FOOT_SWITCH_INPUT_MODE <> INTERN.PREV_SRC_FOOT_SWITCH_INPUT_MODE THEN
			PA.FOOT_SWITCH_INPUT_MODE := INTERN.SRC_FOOT_SWITCH_INPUT_MODE;
		END_IF
		IF INTERN.SRC_LIQUID_LEVEL_INPUT_MODE <> INTERN.PREV_SRC_LIQUID_LEVEL_INPUT_MODE THEN
			PA.LIQUID_LEVEL_INPUT_MODE := INTERN.SRC_LIQUID_LEVEL_INPUT_MODE;
		END_IF
		IF INTERN.SRC_STATE_OUTPUT_MODE <> INTERN.PREV_SRC_STATE_OUTPUT_MODE THEN
			PA.STATE_OUTPUT_MODE := INTERN.SRC_STATE_OUTPUT_MODE;
		END_IF
		IF INTERN.SRC_COMMUNICATION_ADDRESS <> INTERN.PREV_SRC_COMMUNICATION_ADDRESS THEN
			PA.COMMUNICATION_ADDRESS := INTERN.SRC_COMMUNICATION_ADDRESS;
		END_IF
		IF INTERN.SRC_BAUD_RATE_INDEX <> INTERN.PREV_SRC_BAUD_RATE_INDEX THEN
			PA.BAUD_RATE_INDEX := INTERN.SRC_BAUD_RATE_INDEX;
		END_IF
	END_IF

	INTERN.PREV_SRC_MAX_MOTOR_SPEED         := INTERN.SRC_MAX_MOTOR_SPEED;
	INTERN.PREV_SRC_CALIBRATION_COEFFICIENT := INTERN.SRC_CALIBRATION_COEFFICIENT;
	INTERN.PREV_SRC_FOOT_SWITCH_INPUT_MODE  := INTERN.SRC_FOOT_SWITCH_INPUT_MODE;
	INTERN.PREV_SRC_LIQUID_LEVEL_INPUT_MODE := INTERN.SRC_LIQUID_LEVEL_INPUT_MODE;
	INTERN.PREV_SRC_STATE_OUTPUT_MODE       := INTERN.SRC_STATE_OUTPUT_MODE;
	INTERN.PREV_SRC_COMMUNICATION_ADDRESS   := INTERN.SRC_COMMUNICATION_ADDRESS;
	INTERN.PREV_SRC_BAUD_RATE_INDEX         := INTERN.SRC_BAUD_RATE_INDEX;

	//--- Parameters used by the pump : always from PA
	INTERN.CMD_MAX_SPEED      := PA.MAX_MOTOR_SPEED;
	INTERN.CMD_CALIB_COEF     := PA.CALIBRATION_COEFFICIENT;
	INTERN.CMD_FOOT_MODE      := PA.FOOT_SWITCH_INPUT_MODE;
	INTERN.CMD_LEVEL_MODE     := PA.LIQUID_LEVEL_INPUT_MODE;
	INTERN.CMD_STATE_OUT_MODE := PA.STATE_OUTPUT_MODE;
	INTERN.CMD_ADDRESS        := PA.COMMUNICATION_ADDRESS;
	INTERN.CMD_BAUD_INDEX     := PA.BAUD_RATE_INDEX;

	//--- Parameter validity
	INTERN.PARAM_VALID := (WORD_TO_UINT(INTERN.CMD_ADDRESS) >= 1) AND (WORD_TO_UINT(INTERN.CMD_ADDRESS) <= 31)
	                      AND (WORD_TO_UINT(INTERN.CMD_BAUD_INDEX) <= 7)
	                      AND (INTERN.CMD_MAX_SPEED > 0.0) AND (INTERN.CMD_CALIB_COEF > 0.0);

	//--- Flash save : 1 s pulse on rising edge, only with valid parameters
	R_TRIG_FLASH(CLK := INTERN.FLASH_SAVE_REQUEST);
	TP_FLASH(IN := R_TRIG_FLASH.Q AND INTERN.PARAM_VALID, PT := T#1S);
	INTERN.CMD_SAVE_FLASH := TP_FLASH.Q;

	//--- Write triggers (rising edge channels)
	// Square wave 500 ms : each rising edge = one write request
	TON_PULSE(IN := NOT TON_PULSE.Q, PT := T#250MS);
	IF TON_PULSE.Q THEN
		INTERN.PULSE_500MS := NOT INTERN.PULSE_500MS;
	END_IF

	// Command trigger : automatic, 3 s of edges after any command change
	INTERN.CMD_CHANGED := (INTERN.CMD_RUN <> INTERN.PREV_RUN) OR (INTERN.CMD_CLOCKWISE <> INTERN.PREV_CLOCKWISE)
	                      OR (INTERN.CMD_VOLUME_MODE <> INTERN.PREV_VOLUME_MODE) OR (INTERN.CMD_SAVE_FLASH <> INTERN.PREV_SAVE_FLASH)
	                      OR (INTERN.CMD_SPEED <> INTERN.PREV_SPEED) OR (INTERN.CMD_MAX_SPEED <> INTERN.PREV_MAX_SPEED)
	                      OR (INTERN.CMD_RUN_SETPOINT <> INTERN.PREV_RUN_SETPOINT);
	INTERN.PREV_RUN          := INTERN.CMD_RUN;
	INTERN.PREV_CLOCKWISE    := INTERN.CMD_CLOCKWISE;
	INTERN.PREV_VOLUME_MODE  := INTERN.CMD_VOLUME_MODE;
	INTERN.PREV_SAVE_FLASH   := INTERN.CMD_SAVE_FLASH;
	INTERN.PREV_SPEED        := INTERN.CMD_SPEED;
	INTERN.PREV_MAX_SPEED    := INTERN.CMD_MAX_SPEED;
	INTERN.PREV_RUN_SETPOINT := INTERN.CMD_RUN_SETPOINT;

	TOF_CMD_WINDOW(IN := INTERN.CMD_CHANGED, PT := T#3S);
	INTERN.CMD_WINDOW  := TOF_CMD_WINDOW.Q;
	INTERN.CMD_TRIGGER := INTERN.CMD_WINDOW AND (INTERN.CMD_MAX_SPEED > 0.0) AND INTERN.PULSE_500MS;

	// Configuration trigger : only while writing is enabled and parameters are valid
	INTERN.CONFIG_TRIGGER := INTERN.PARAM_WRITE_ENABLE AND INTERN.PARAM_VALID AND INTERN.PULSE_500MS;


//------------------------------------------------------------------------------
// 3. OUTPUTS
//------------------------------------------------------------------------------
	//--- COM : control mode status to SCADA, HMI and WEBVISU
	COM.SCADA_OUTPUT_LOCAL_FUXA_ACTIVE := INTERN.LOCAL_FUXA;
	COM.SCADA_OUTPUT_LOCAL_HMI_ACTIVE  := INTERN.LOCAL_HMI;
	COM.HMI_OUTPUT_LOCAL_ACTIVE        := INTERN.LOCAL_HMI;
	COM.WEBVISU_OUTPUT_LOCAL_ACTIVE        := INTERN.LOCAL_WEBVISU;
	COM.WEBVISU_OUTPUT_LOCAL_HMI_ACTIVE  := INTERN.LOCAL_HMI;
	COM.WEBVISU_OUTPUT_LOCAL_FUXA_ACTIVE := INTERN.LOCAL_FUXA;

	//--- COM : Modbus RTU coils
	COM.COM_OUTPUT_COILS[0] := INTERN.CMD_RUN;           // 0x0001
	COM.COM_OUTPUT_COILS[1] := INTERN.CMD_CLOCKWISE;     // 0x0002
	COM.COM_OUTPUT_COILS[2] := INTERN.CMD_SAVE_FLASH;    // 0x0003
	COM.COM_OUTPUT_COILS[3] := INTERN.CMD_VOLUME_MODE;   // 0x0004

	//--- COM : Modbus RTU holding registers and write triggers
	// Command registers 0x4001..0x4006 (sent on the command trigger)
	FNC_REAL_TO_WORDS(Real_value := INTERN.CMD_SPEED,     High_word => COM.COM_OUTPUT_HR_CMD[1], Low_word => COM.COM_OUTPUT_HR_CMD[0]);   // 0x4001-4002
	FNC_REAL_TO_WORDS(Real_value := INTERN.CMD_MAX_SPEED, High_word => COM.COM_OUTPUT_HR_CMD[3], Low_word => COM.COM_OUTPUT_HR_CMD[2]);   // 0x4003-4004
	IF INTERN.CMD_VOLUME_MODE THEN
		// Run setpoint 0x4005-4006, volume mode : 32-bit REAL (ml)
		FNC_REAL_TO_WORDS(Real_value := INTERN.CMD_RUN_SETPOINT, High_word => COM.COM_OUTPUT_HR_CMD[5], Low_word => COM.COM_OUTPUT_HR_CMD[4]);
	ELSE
		// Run setpoint 0x4005-4006, time mode : 32-bit UDINT (ms)
		INTERN.UDINT_TEMP        := REAL_TO_UDINT(MAX(INTERN.CMD_RUN_SETPOINT, 0.0));
		COM.COM_OUTPUT_HR_CMD[4] := UDINT_TO_WORD(INTERN.UDINT_TEMP);
		COM.COM_OUTPUT_HR_CMD[5] := UDINT_TO_WORD(SHR(INTERN.UDINT_TEMP, 16));
	END_IF

	// Configuration registers 0x400B..0x4011 (sent on the configuration trigger), updated only while enabled and valid
	IF INTERN.PARAM_WRITE_ENABLE AND INTERN.PARAM_VALID THEN
		FNC_REAL_TO_WORDS(Real_value := INTERN.CMD_CALIB_COEF, High_word => COM.COM_OUTPUT_HR_CONFIG[1], Low_word => COM.COM_OUTPUT_HR_CONFIG[0]);   // 0x400B-400C
		COM.COM_OUTPUT_HR_CONFIG[2] := INTERN.CMD_FOOT_MODE;        // 0x400D
		COM.COM_OUTPUT_HR_CONFIG[3] := INTERN.CMD_LEVEL_MODE;       // 0x400E
		COM.COM_OUTPUT_HR_CONFIG[4] := INTERN.CMD_STATE_OUT_MODE;   // 0x400F
		COM.COM_OUTPUT_HR_CONFIG[5] := INTERN.CMD_ADDRESS;          // 0x4010
		COM.COM_OUTPUT_HR_CONFIG[6] := INTERN.CMD_BAUD_INDEX;       // 0x4011
	END_IF

	// Write triggers
	COM.COM_OUTPUT_CMD_TRIGGER    := INTERN.CMD_TRIGGER;
	COM.COM_OUTPUT_CONFIG_TRIGGER := INTERN.CONFIG_TRIGGER;

	//--- COM : feedback to SCADA, HMI and WEBVISU
	COM.SCADA_OUTPUT_FIRMWARE_VERSION                          := INTERN.FBK_FIRMWARE_VERSION;
	COM.HMI_OUTPUT_FIRMWARE_VERSION                            := INTERN.FBK_FIRMWARE_VERSION;
	COM.WEBVISU_OUTPUT_FIRMWARE_VERSION                            := INTERN.FBK_FIRMWARE_VERSION;
	COM.SCADA_OUTPUT_HARDWARE_VERSION                          := INTERN.FBK_HARDWARE_VERSION;
	COM.HMI_OUTPUT_HARDWARE_VERSION                            := INTERN.FBK_HARDWARE_VERSION;
	COM.WEBVISU_OUTPUT_HARDWARE_VERSION                            := INTERN.FBK_HARDWARE_VERSION;
	COM.SCADA_OUTPUT_TEMPERATURE                               := INTERN.FBK_TEMPERATURE;
	COM.HMI_OUTPUT_TEMPERATURE                                 := INTERN.FBK_TEMPERATURE;
	COM.WEBVISU_OUTPUT_TEMPERATURE                                 := INTERN.FBK_TEMPERATURE;
	COM.SCADA_OUTPUT_FLOAT_LEVEL_ALARM                         := INTERN.FBK_LEVEL_ALARM;
	COM.HMI_OUTPUT_FLOAT_LEVEL_ALARM                           := INTERN.FBK_LEVEL_ALARM;
	COM.WEBVISU_OUTPUT_FLOAT_LEVEL_ALARM                           := INTERN.FBK_LEVEL_ALARM;
	COM.SCADA_OUTPUT_DIGITAL_OUTPUT_VALUE                      := INTERN.FBK_DIGITAL_OUTPUT;
	COM.HMI_OUTPUT_DIGITAL_OUTPUT_VALUE                        := INTERN.FBK_DIGITAL_OUTPUT;
	COM.WEBVISU_OUTPUT_DIGITAL_OUTPUT_VALUE                        := INTERN.FBK_DIGITAL_OUTPUT;
	COM.SCADA_OUTPUT_REAL_TIME_RUN_TIME_OR_VOLUME.Real_value   := INTERN.FBK_RUN_ACTUAL;
	COM.HMI_OUTPUT_REAL_TIME_RUN_TIME_OR_VOLUME.Real_value     := INTERN.FBK_RUN_ACTUAL;
	COM.WEBVISU_OUTPUT_REAL_TIME_RUN_TIME_OR_VOLUME.Real_value     := INTERN.FBK_RUN_ACTUAL;
	COM.SCADA_OUTPUT_ACCUMULATED_RUN_TIME_OR_VOLUME.Real_value := INTERN.FBK_RUN_TOTAL;
	COM.HMI_OUTPUT_ACCUMULATED_RUN_TIME_OR_VOLUME.Real_value   := INTERN.FBK_RUN_TOTAL;
	COM.WEBVISU_OUTPUT_ACCUMULATED_RUN_TIME_OR_VOLUME.Real_value   := INTERN.FBK_RUN_TOTAL;


                
END_FUNCTION_BLOCK

FUNCTION FNC_REAL_TO_WORDS : BOOL
  VAR_INPUT
    Real_value : REAL;  (* Value to split *)
  END_VAR
  VAR_OUTPUT
    High_word : WORD;  (* Most significant word *)
    Low_word : WORD;  (* Least significant word *)
  END_VAR
  VAR
    Conversion : DUT_Union_Real_Word;  (* REAL / 2 WORD overlay *)
  END_VAR

                  
//==============================================================================
// FNC_REAL_TO_WORDS
// REAL (IEEE 754) -> two Modbus words
// Call: FNC_REAL_TO_WORDS(Real_value := x, High_word => ..., Low_word => ...);
//==============================================================================

Conversion.Real_value := Real_value;
Low_word  := Conversion.Word_value[0];
High_word := Conversion.Word_value[1];
FNC_REAL_TO_WORDS := TRUE;

                
END_FUNCTION

FUNCTION FNC_WORDS_TO_REAL : REAL
  VAR_INPUT
    High_word : WORD;  (* Most significant word *)
    Low_word : WORD;  (* Least significant word *)
  END_VAR
  VAR
    Conversion : DUT_Union_Real_Word;  (* REAL / 2 WORD overlay *)
  END_VAR

                  
//==============================================================================
// FNC_WORDS_TO_REAL
// Two Modbus words -> REAL (IEEE 754)
// ABCD device: High_word = lower address, CDAB device: Low_word = lower address
//==============================================================================

Conversion.Word_value[0] := Low_word;
Conversion.Word_value[1] := High_word;
FNC_WORDS_TO_REAL := Conversion.Real_value;

                
END_FUNCTION

FUNCTION GFC_COM_IN : BOOL

                  
//==============================================================================
// GFC_COM_IN
// Modbus (GVL_MODBUS) -> GVL_COM : RTU equipment, SCADA FUXA, HMI
// Simple copies only, no conversion (conversions are done in the FBs)
//==============================================================================

//------------------------------------------------------------------------------
// COM : Modbus RTU, from equipment
//------------------------------------------------------------------------------
	//--- ADM100W_1
	GVL_COM.COM_ADM100W_1.COM_INPUT_IR    := GVL_MODBUS.ADM100W_InputRegisters;   // Input registers 0..87
	GVL_COM.COM_ADM100W_1.COM_INPUT_COILS := GVL_MODBUS.ADM100W_Alarms;           // Coils 0..9 (alarms)

	//--- DIP1500_1
	GVL_COM.COM_DIP1500_1.COM_INPUT_IR          := GVL_MODBUS.DIP1500_InputRegisters;     // Input registers 0x3001..0x3005
	GVL_COM.COM_DIP1500_1.COM_INPUT_HR_COUNTERS := GVL_MODBUS.DIP1500_Holding_Counters;   // Holding registers 0x4007..0x400A


//------------------------------------------------------------------------------
// SCADA FUXA : coils (FUXA 000001...)
//------------------------------------------------------------------------------
	//--- DOSENSOR_1
	GVL_COM.COM_DOSENSOR_1.SCADA_INPUT_CALIBRATION_HIGH := GVL_MODBUS.Coils_TCP_HMI[0].0;   // 1 | DO Calibration High
	GVL_COM.COM_DOSENSOR_1.SCADA_INPUT_CALIBRATION_LOW  := GVL_MODBUS.Coils_TCP_HMI[0].1;   // 2 | DO Calibration Low
	GVL_COM.COM_DOSENSOR_1.SCADA_INPUT_LOCAL_REQUEST    := GVL_MODBUS.Coils_TCP_HMI[0].7;   // 8 | DO Sensor Local Request
	GVL_COM.COM_DOSENSOR_1.SCADA_INPUT_AUTO_REQUEST     := GVL_MODBUS.Coils_TCP_HMI[1].0;   // 9 | DO Sensor Auto Request

	//--- DIP1500_1
	GVL_COM.COM_DIP1500_1.SCADA_INPUT_MOTOR_START_STOP   := GVL_MODBUS.Coils_TCP_HMI[0].2;   // 3 | DIP1500 Motor Start Stop
	GVL_COM.COM_DIP1500_1.SCADA_INPUT_MOTOR_DIRECTION    := GVL_MODBUS.Coils_TCP_HMI[0].3;   // 4 | DIP1500 Motor Direction
	GVL_COM.COM_DIP1500_1.SCADA_INPUT_FLASH_SAVE         := GVL_MODBUS.Coils_TCP_HMI[0].4;   // 5 | DIP1500 Flash Save
	GVL_COM.COM_DIP1500_1.SCADA_INPUT_OPERATION_MODE     := GVL_MODBUS.Coils_TCP_HMI[0].5;   // 6 | DIP1500 Operation Mode
	GVL_COM.COM_DIP1500_1.SCADA_INPUT_PARAM_WRITE_ENABLE := GVL_MODBUS.Coils_TCP_HMI[0].6;   // 7 | DIP1500 Parameter Write Enable
	GVL_COM.COM_DIP1500_1.SCADA_INPUT_LOCAL_REQUEST      := GVL_MODBUS.Coils_TCP_HMI[1].1;   // 10 | DIP1500 Local Request
	GVL_COM.COM_DIP1500_1.SCADA_INPUT_AUTO_REQUEST       := GVL_MODBUS.Coils_TCP_HMI[1].2;   // 11 | DIP1500 Auto Request

	//--- ADM100W_1
	GVL_COM.COM_ADM100W_1.SCADA_INPUT_LOCAL_REQUEST := GVL_MODBUS.Coils_TCP_HMI[1].3;   // 12 | ADM100W Local Request
	GVL_COM.COM_ADM100W_1.SCADA_INPUT_AUTO_REQUEST  := GVL_MODBUS.Coils_TCP_HMI[1].4;   // 13 | ADM100W Auto Request

	//--- UPI_LOCAL_FUXA
	GVL_COM.COM_UPI_LOCAL_FUXA.SCADA_INPUT_LOCAL_REQUEST := GVL_MODBUS.Coils_TCP_HMI[1].5;   // 14 | Global Local FUXA Request
	GVL_COM.COM_UPI_LOCAL_FUXA.SCADA_INPUT_AUTO_REQUEST  := GVL_MODBUS.Coils_TCP_HMI[1].6;   // 15 | Global Auto FUXA Request


